(* CODESYS project process.library
   DefaultNamespace: KOSTAL.AF2024.Core.Process
   DocFormat: reStructuredText
   Description: Core Functionalities UTF16
   Author: Frank Dümpelmann
   Title: KOSTAL.AF2024.Core.Process
   Version: 1.0.999.1
   Company: KOSTAL GmbH & Co.KG
   Placeholder: KOSTAL.AF2024.Core.Process

Project tree, tasks and I/O mapping:
  libraries: KOSTAL.AF2024.Core.functionResponse, 1.0.0.0 (KOSTAL GmbH & Co.KG); KOSTAL.AF2024.Core.ListOf, 1.0.0.0 (KOSTAL GmbH & Co.KG); KOSTAL.AF2024.Core.Settings, 1.0.0.0 (KOSTAL GmbH & Co.KG); KOSTAL.AF2024.Core.StringTools, 1.0.0.0 (KOSTAL GmbH & Co.KG); KOSTAL.AF2024.Core.System, 1.0.0.0 (KOSTAL GmbH & Co.KG)
  _Global/
    E_/
      data type E_PROCESS_CONDITION_DEFAULT_PRIORITYLEVEL
  Condition/
    function block FB_processCondition [ST]: clear, CopyFrom, CopyTo, FB_init, getPriority, isActive, isError, isFail, isInfo, isMasterMessage, isMessage, isPass, isText, Message, Message_Owner, PriorityLevel_Error, PriorityLevel_Info, PriorityLevel_MasterMessage, PriorityLevel_Message, PriorityLevel_Text, setMessage, setMessageFail, setMessagePass
    interface I_processCondition: CopyTo, getPriority, isActive, isError, isFail, isInfo, isMasterMessage, isMessage, isPass, isText, Message, PriorityLevel_Error, PriorityLevel_Info, PriorityLevel_MasterMessage, PriorityLevel_Message, PriorityLevel_Text
    interface I_processCondition_CopyFrom: CopyFrom
    interface I_processCondition_Owner: clear, CopyFrom, CopyTo, getPriority, isActive, isError, isFail, isInfo, isMasterMessage, isMessage, isPass, isText, Message, Message_Owner, PriorityLevel_Error, PriorityLevel_Info, PriorityLevel_MasterMessage, PriorityLevel_Message, PriorityLevel_Text, setMessage, setMessageFail, setMessagePass
  DeviceState/
    interface I_T_deviceState: Fault, Off, On, Operational
    interface I_T_deviceState_Owner: ClearPlcState, Fault, Off, On, Operational
    function block T_deviceState [ST]: Clear, ClearPlcState, CopyFrom, CopyTo, Fault, Off, On, Operational
  Message/
    messageText/
      interface I_T_messageText: CopyTo, line_01, toString
      interface I_T_messageText_CopyFrom: CopyFrom
      interface I_T_messageText_Owner: clear, CopyFrom, CopyTo, line_01, toString
      function block T_messageText [ST]: clear, CopyFrom, CopyTo, line_01, toString
    messageText_2_lines/
      interface I_T_messageText_2_lines: line_02
      interface I_T_messageText_2_lines_Owner: line_02
      function block T_messageText_2_lines [ST]: clear, CopyFrom, line_02, toString
    messageText_3_lines/
      interface I_T_messageText_3_lines: line_03
      interface I_T_messageText_3_lines_Owner: line_03
      function block T_messageText_3_lines [ST]: clear, CopyFrom, line_03, toString
  PlcState/
    interface I_T_plcState: busy, CopyTo, description, fail, finish, pass, ready
    interface I_T_plcState_CopyFrom: CopyFrom
    interface I_T_plcState_Owner: busy, clear, CopyFrom, CopyTo, description, fail, finish, pass, ready
    function block T_plcState [ST]: busy, clear, CopyFrom, CopyTo, description, fail, finish, pass, ready
  ProcessMode/
    interface I_T_processMode: automatic, CopyTo, manual
    interface I_T_processMode_CopyFrom: CopyFrom
    interface I_T_processMode_Owner: automatic, clear, CopyFrom, CopyTo, manual
    function block T_processMode [ST]: automatic, clear, CopyFrom, CopyTo, manual
  Project Information/
    function F_GetCompany [ST]
    function F_GetTitle [ST]
    function F_GetVersion [ST]
  Step/
    GVL/
      global variables ProcessStep_GVL
    processStep/
      function block FB_processStep [ST]: actual, clear, CopyFrom, CopyTo, DEC, Header, INC, init, request, set, toggle
      interface I_processStep: actual, CopyTo, request, toggle
      interface I_processStep_CopyFrom: CopyFrom
      interface I_processStep_Owner: actual, clear, CopyFrom, CopyTo, DEC, Header, INC, init, request, set, toggle
    processStep_Control/
      StepMemory/
        ListOf/
          function block FB_ListOf_T_StepMemory [ST]: _get_I, _get_I_RO, _removePayLoad, _verifyMember, Add_DUT, Clear, CopyFrom, CopyTo, Delete_DUT, Get_I, Get_I_RO, MaxEntries, NumberOfMember
          interface I_ListOf_StepMemory: Add_DUT, Clear, CopyFrom, CopyTo, Delete_DUT, Get_I, Get_I_RO, MaxEntries, NumberOfMember
          interface I_ListOf_StepMemory_CopyFrom: CopyFrom
          interface I_ListOf_StepMemory_RO: CopyTo, Get_I_RO, MaxEntries, NumberOfMember
        interface I_T_StepMemory: Clear, CopyFrom, Actual, RegKey, Request
        interface I_T_StepMemory_CopyFrom: CopyFrom
        interface I_T_StepMemory_RO: CopyTo, Actual, RegKey, Request
        function block T_StepMemory [ST]: Clear, CopyFrom, CopyTo, Actual, RegKey, Request
      function block FB_ProcessStep_Control [ST]: FB_exit, FB_init, _DEC, _INC, _init, _set, _modeAutomatik, _backward, _forward, _modeManual, _addStep, _removeStep, _preset, DEC, INC, init, set, Control, clear, CopyFrom, Header, LinkManual, BackwardDone, Done, FromBackStep, LastUsedKey, StepMemory, StepMemory_RO, StepNumberHome, Condition, DisableBackward, JumpAddress, ManualWithCondition, mode
      interface I_ProcessStep_Control: BackwardDone, Done, FromBackStep, LastUsedKey, StepMemory_RO, StepNumberHome, Condition, DisableBackward, JumpAddress, ManualWithCondition, mode
      interface I_ProcessStep_Control_Owner: Control, Header, LinkManual, BackwardDone, Done, FromBackStep, LastUsedKey, StepMemory, StepMemory_RO, StepNumberHome, Condition, DisableBackward, JumpAddress, ManualWithCondition, mode
    processStep_Flow/
      function block FB_processStep_Flow [ST]: clear, Header, init, isActive, isCalledExternally, NotFound
      interface I_processStep_Flow: isCalledExternally, NotFound
      interface I_processStep_Flow_Owner: clear, Header, init, isActive, isCalledExternally, NotFound
  Version/
    global variables Global_Version
*)

// _Global/E_/E_PROCESS_CONDITION_DEFAULT_PRIORITYLEVEL
(*
Description
===========
| Levels of message priorities
| Intermediate values can be used to overrule other messages of the same level
| 1..999: INFORMATION - Display less important information (Color: grey)
| 1000..1999: TEXT_ONLY - To display information (Color: green)
| 2000..2999: MESSAGE - Order to the operator, e.g. 'Insert part' (Color: blue)
| 3000..3999: MASTERMESSAGE - Message to be displayed in upper HMI levels (Color: blue)
| 4000..4999: ERROR - Error message (Color: orange)

*)

{attribute 'qualified_only'}
TYPE E_PROCESS_CONDITION_DEFAULT_PRIORITYLEVEL :
(
	NONE 			:= 0,
	INFORMATION		:= 1,
	TEXT_ONLY		:= 1000,
	MESSAGE			:= 2000,
	MASTERMESSAGE	:= 3000,
	ERROR			:= 4000
);
END_TYPE

// Step/GVL/ProcessStep_GVL
{attribute 'qualified_only'}
VAR_GLOBAL CONSTANT
	PROCESS_STEP_INITIALIZE_STEP	: INT:= INT#32767; //INT[max] 16#7FFF;
END_VAR

// Version/Global_Version
{attribute 'TcGenerated'}
{attribute 'no-analysis'}
{attribute 'linkalways'}
// This function has been automatically generated from the project information.
VAR_GLOBAL CONSTANT
	{attribute 'const_non_replaced'}
	stLibVersion_KOSTAL_AF2024_Core_Process : ST_LibVersion := (iMajor := 1, iMinor := 0, iBuild := 999, iRevision := 1, nFlags := 1, sVersion := '1.0.999.1');
END_VAR

// Condition/FB_processCondition
(*

:Author: Frank Dümpelmann <f.duempelmann@kostal.com>
:Date: 2018-10-26

Function
========
| Data structure representing the status of users/stations 
| Used for communication to superior instances, e.g. HMI

Usage notes
===============
| Call method setMessage from User/Station to set Message Text and priority level
| Call methods is... from the superior instance to get the user's status 
| Read message text from property message 

Methods and Properties
======================
| See bottom of this document for a detailed description of each method or property
*)

{attribute 'enable_dynamic_creation'}
FUNCTION_BLOCK PUBLIC FB_processCondition IMPLEMENTS I_processCondition, I_processCondition_CopyFrom, I_processCondition_Owner

VAR
	_priority	: INT;	//Priority of message
	
	_message	: T_messageText_3_lines;
	
	_pass		: BOOL;
	_fail		: BOOL;
END_VAR

(*
Description
===========
| Clears existing message
*)

METHOD PUBLIC clear

_priority:= E_PROCESS_CONDITION_DEFAULT_PRIORITYLEVEL.NONE;

_message.clear();
_pass := _fail := false;
END_METHOD

METHOD PUBLIC CopyFrom : BOOL
VAR_INPUT
	IN	: KOSTAL_AF2024_Core_System.I_Interface;
END_VAR

VAR
	_obj		: I_processCondition;
	_obj2		: I_processCondition_Owner;
	_bFound	:	BOOL;
END_VAR

IF IN = 0 THEN	RETURN;	END_IF

clear();

//-----------------------------------------

_bFound:= __QUERYINTERFACE(IN, _obj);

IF _bFound AND_THEN _obj <> 0 THEN
	
	_priority:= _obj.getPriority();
	
	_message.CopyFrom(_obj.Message);
	
	_pass := _obj.isPass();
	_fail := _obj.isFail();
	
	
	CopyFrom:= TRUE;
	
	RETURN;
	
END_IF

//-----------------------------------------

_bFound:= __QUERYINTERFACE(IN, _obj2);

IF _bFound AND_THEN _obj2 <> 0 THEN
	
	_priority:= _obj2.getPriority();
	
	_message.CopyFrom(_obj2.Message);
	
	_pass := _obj2.isPass();
	_fail := _obj2.isFail();
	
	CopyFrom:= TRUE;

	RETURN;
	
END_IF
END_METHOD

METHOD PUBLIC CopyTo : BOOL
VAR_INPUT
	IN	:	I_processCondition_CopyFrom;
END_VAR

IF IN = 0 THEN	RETURN;	END_IF

CopyTo:= IN.CopyFrom(THIS^);
END_METHOD

(*
Description
===========
| To be called automatically!
*)
METHOD FB_init : BOOL
VAR_INPUT
	bInitRetains : BOOL; // if TRUE, the retain variables are initialized (warm start / cold start)
	bInCopyCode : BOOL;  // if TRUE, the instance afterwards gets moved into the copy code (online change)
END_VAR
//_infoPriorityLevel			:= E_PROCESS_CONDITION_DEFAULT_PRIORITYLEVEL.INFORMATION; 
//_textPriorityLevel			:= E_PROCESS_CONDITION_DEFAULT_PRIORITYLEVEL.TEXT_ONLY;		//define the priority level from which priority a message is an user relative text 
//_messagePriorityLevel		:= E_PROCESS_CONDITION_DEFAULT_PRIORITYLEVEL.MESSAGE;		//define the priority level from which priority a message is an user relative message 
//_masterMessagePriorityLevel	:= E_PROCESS_CONDITION_DEFAULT_PRIORITYLEVEL.MASTERMESSAGE;	//define the priority level from which priority a message is an user relative error 
//_errorPriorityLevel			:= E_PROCESS_CONDITION_DEFAULT_PRIORITYLEVEL.ERROR;			//define the priority level from which priority a message is an user relative error
END_METHOD

METHOD PUBLIC getPriority : INT
VAR_INPUT
END_VAR

getPriority:= _priority;
END_METHOD

(*
Description
===========
| Returns TRUE if the user has a text, message or error to display
*)

METHOD PUBLIC isActive : BOOL
VAR_INPUT
END_VAR

isActive:= _priority <> E_PROCESS_CONDITION_DEFAULT_PRIORITYLEVEL.NONE;
END_METHOD

(*
Description
===========
| Returns TRUE if the user has an error to display
*)
METHOD PUBLIC isError : BOOL
VAR_INPUT
END_VAR

isError:= _priority >= E_PROCESS_CONDITION_DEFAULT_PRIORITYLEVEL.ERROR;
END_METHOD

METHOD PUBLIC isFail : BOOL
VAR_INPUT
END_VAR
isFail := (isMessage() OR isMasterMessage()) AND _fail;
END_METHOD

(*
Description
===========
| Returns TRUE if the user has a message to display
*)
METHOD PUBLIC isInfo : BOOL
VAR_INPUT
END_VAR

isInfo:= (_priority >= E_PROCESS_CONDITION_DEFAULT_PRIORITYLEVEL.INFORMATION) AND (_priority < E_PROCESS_CONDITION_DEFAULT_PRIORITYLEVEL.TEXT_ONLY);
END_METHOD

(*
Description
===========
| Returns TRUE if the user has a master message to display
*)
METHOD PUBLIC isMasterMessage : BOOL
VAR_INPUT
END_VAR

isMasterMessage:= (_priority >= E_PROCESS_CONDITION_DEFAULT_PRIORITYLEVEL.MASTERMESSAGE) AND (_priority < E_PROCESS_CONDITION_DEFAULT_PRIORITYLEVEL.ERROR);
END_METHOD

(*
Description
===========
| Returns TRUE if the user has a message to display
*)
METHOD PUBLIC isMessage : BOOL
VAR_INPUT
END_VAR

isMessage:= (_priority >= E_PROCESS_CONDITION_DEFAULT_PRIORITYLEVEL.MESSAGE) AND (_priority < E_PROCESS_CONDITION_DEFAULT_PRIORITYLEVEL.MASTERMESSAGE);
END_METHOD

METHOD PUBLIC isPass : BOOL
VAR_INPUT
END_VAR
isPass := (isMessage() OR isMasterMessage()) AND _pass;
END_METHOD

(*
Description
===========
| Returns TRUE if the user has a text to display
*)
METHOD PUBLIC isText : BOOL

isText:= (_priority >= E_PROCESS_CONDITION_DEFAULT_PRIORITYLEVEL.TEXT_ONLY) AND (_priority < E_PROCESS_CONDITION_DEFAULT_PRIORITYLEVEL.MESSAGE);
END_METHOD

(*
Description
===========
| Message to display in three lines
*)

PROPERTY PUBLIC Message : I_T_messageText_3_lines
GET


Message := _message;
END_GET
END_PROPERTY

(*
Description
===========
| Message to display in three lines
*)

PROPERTY PUBLIC Message_Owner : I_T_messageText_3_lines_Owner
GET


Message_Owner := _message;
END_GET
END_PROPERTY

PROPERTY PUBLIC PriorityLevel_Error : INT
GET

PriorityLevel_Error := E_PROCESS_CONDITION_DEFAULT_PRIORITYLEVEL.ERROR;// _errorPriorityLevel;
END_GET
END_PROPERTY

PROPERTY PUBLIC PriorityLevel_Info : INT
GET

PriorityLevel_Info := E_PROCESS_CONDITION_DEFAULT_PRIORITYLEVEL.INFORMATION;
END_GET
END_PROPERTY

PROPERTY PUBLIC PriorityLevel_MasterMessage : INT
GET

PriorityLevel_MasterMessage := E_PROCESS_CONDITION_DEFAULT_PRIORITYLEVEL.MASTERMESSAGE;
END_GET
END_PROPERTY

PROPERTY PUBLIC PriorityLevel_Message : INT
GET

PriorityLevel_Message := E_PROCESS_CONDITION_DEFAULT_PRIORITYLEVEL.MESSAGE;
END_GET
END_PROPERTY

PROPERTY PUBLIC PriorityLevel_Text : INT
GET

PriorityLevel_Text := E_PROCESS_CONDITION_DEFAULT_PRIORITYLEVEL.TEXT_ONLY;
END_GET
END_PROPERTY

(*
Description
===========
| Sets message text and priority level for the user, in case the priority is higher than the existing message's priority 
| Existing messages with the same or lower priority are cleared
| Parameters:
| 	priority: INT - See E_PROCESS_CONDITION_DEFAULT_PRIORITYLEVEL for a detailed description
|	message: FB_messageText_3_lines - Content of the message
| Return value:
| 	FB_functionResponse: 
|		result: BOOL - Message ist set (no existing message with higher priority)
|		status: STRING(255) - Error description
*)

METHOD PUBLIC setMessage : KOSTAL_AF2024_Core_functionResponse.T_functionResponse

VAR_INPUT
	priority	: INT;
	message		: I_T_messageText_3_lines;
END_VAR
IF message = 0 THEN 
	setMessage.Status	:= "Message is invalid";
	setMessage.Success	:= FALSE;
	RETURN;	
END_IF

IF priority > _priority THEN
	setMessage.clear();
	_priority	:= priority;
	_message.CopyFrom(message);
	_pass := FALSE;
	_fail := FALSE;
	setMessage.Success	:= TRUE;

ELSE

	setMessage.Status	:= "actual priority is higher";
	setMessage.Success	:= FALSE;

END_IF
END_METHOD

(*
Description
===========
| Sets message text and priority level for the user, in case the priority is higher than the existing message's priority  
| Message is displayed as "Fail" (red) in WInHMI
| Existing messages with the same or lower priority are cleared
| Parameters:
| 	priority: INT - See E_PROCESS_CONDITION_DEFAULT_PRIORITYLEVEL for a detailed description
|	message: FB_messageText_3_lines - Content of the message
| Return value:
| 	FB_functionResponse: 
|		result: BOOL - Message ist set (no existing message with higher priority)
|		status: STRING(255) - Error description
*)

METHOD PUBLIC setMessageFail : KOSTAL_AF2024_Core_functionResponse.T_functionResponse

VAR_INPUT
	priority	: INT;
	message		: I_T_messageText_3_lines;
END_VAR
IF message = 0 THEN 
	setMessageFail.Status	:= "Message is invalid";
	setMessageFail.Success	:= FALSE;
	RETURN;	
END_IF

IF priority > _priority THEN
	setMessageFail.clear();
	_priority	:= priority;
	_message.CopyFrom(message);
	_pass := FALSE;
	_fail := TRUE;
	
	setMessageFail.Success	:= TRUE;

ELSE

	setMessageFail.Status	:= "actual priority is higher";
	setMessageFail.Success	:= FALSE;

END_IF
END_METHOD

(*
Description
===========
| Sets message text and priority level for the user, in case the priority is higher than the existing message's priority 
| Message is displayed as "Pass" (green) in WinHMI
| Existing messages with the same or lower priority are cleared
| Parameters:
| 	priority: INT - See E_PROCESS_CONDITION_DEFAULT_PRIORITYLEVEL for a detailed description
|	message: FB_messageText_3_lines - Content of the message
| Return value:
| 	FB_functionResponse: 
|		result: BOOL - Message ist set (no existing message with higher priority)
|		status: STRING(255) - Error description
*)

METHOD PUBLIC setMessagePass : KOSTAL_AF2024_Core_functionResponse.T_functionResponse

VAR_INPUT
	priority	: INT;
	message		: I_T_messageText_3_lines;
END_VAR
IF message = 0 THEN 
	setMessagePass.Status	:= "Message is invalid";
	setMessagePass.Success	:= FALSE;
	RETURN;	
END_IF

IF priority > _priority THEN
	setMessagePass.clear();
	_priority	:= priority;
	_message.CopyFrom(message);
	_pass := TRUE;
	_fail := FALSE;
	
	setMessagePass.Success	:= TRUE;

ELSE

	setMessagePass.Status	:= "actual priority is higher";
	setMessagePass.Success	:= FALSE;

END_IF
END_METHOD

END_FUNCTION_BLOCK

// Condition/I_processCondition
INTERFACE I_processCondition EXTENDS KOSTAL_AF2024_Core_System.I_Interface

METHOD PUBLIC CopyTo : BOOL
VAR_INPUT
	IN	:	I_processCondition_CopyFrom;
END_VAR
END_METHOD

METHOD PUBLIC getPriority : INT
VAR_INPUT
END_VAR
END_METHOD

(*
Description
===========
| Returns TRUE if the user has a text, message or error to display
*)

METHOD PUBLIC isActive : BOOL
VAR_INPUT
END_VAR
END_METHOD

(*
Description
===========
| Returns TRUE if the user has an error to display
*)
METHOD PUBLIC isError : BOOL
VAR_INPUT
END_VAR
END_METHOD

METHOD PUBLIC isFail : BOOL
VAR_INPUT
END_VAR
END_METHOD

(*
Description
===========
| Returns TRUE if the user has a message to display
*)
METHOD PUBLIC isInfo : BOOL
VAR_INPUT
END_VAR
END_METHOD

(*
Description
===========
| Returns TRUE if the user has a master message to display
*)
METHOD PUBLIC isMasterMessage : BOOL
VAR_INPUT
END_VAR
END_METHOD

(*
Description
===========
| Returns TRUE if the user has a message to display
*)
METHOD PUBLIC isMessage : BOOL
VAR_INPUT
END_VAR
END_METHOD

METHOD PUBLIC isPass : BOOL
VAR_INPUT
END_VAR
END_METHOD

(*
Description
===========
| Returns TRUE if the user has a text to display
*)
METHOD PUBLIC isText : BOOL
END_METHOD

(*
Description
===========
| Message to display in three lines
*)

PROPERTY PUBLIC Message : I_T_messageText_3_lines
GET
END_GET
END_PROPERTY

PROPERTY PUBLIC PriorityLevel_Error : INT
GET
END_GET
END_PROPERTY

PROPERTY PUBLIC PriorityLevel_Info : INT
GET
END_GET
END_PROPERTY

PROPERTY PUBLIC PriorityLevel_MasterMessage : INT
GET
END_GET
END_PROPERTY

PROPERTY PUBLIC PriorityLevel_Message : INT
GET
END_GET
END_PROPERTY

PROPERTY PUBLIC PriorityLevel_Text : INT
GET
END_GET
END_PROPERTY

END_INTERFACE

// Condition/I_processCondition_CopyFrom
INTERFACE I_processCondition_CopyFrom EXTENDS KOSTAL_AF2024_Core_System.I_Interface

METHOD PUBLIC CopyFrom : BOOL
VAR_INPUT
	IN	: KOSTAL_AF2024_Core_System.I_Interface;
END_VAR
END_METHOD

END_INTERFACE

// Message/messageText_3_lines/I_T_messageText_3_lines
INTERFACE I_T_messageText_3_lines EXTENDS I_T_messageText_2_lines

PROPERTY PUBLIC line_03 : KOSTAL_AF2024_Core_Settings.T_MaxString
GET
END_GET
END_PROPERTY

END_INTERFACE

// Message/messageText_2_lines/I_T_messageText_2_lines
INTERFACE I_T_messageText_2_lines EXTENDS I_T_messageText

PROPERTY PUBLIC line_02 : KOSTAL_AF2024_Core_Settings.T_MaxString
GET
END_GET
END_PROPERTY

END_INTERFACE

// Message/messageText/I_T_messageText
INTERFACE I_T_messageText EXTENDS KOSTAL_AF2024_Core_System.I_Interface

METHOD PUBLIC CopyTo : bool
VAR_INPUT
	IN	:	I_T_messageText_CopyFrom;
END_VAR
END_METHOD

PROPERTY PUBLIC line_01 : KOSTAL_AF2024_Core_Settings.T_MaxString
GET
END_GET
END_PROPERTY

METHOD PUBLIC toString : KOSTAL_AF2024_Core_Settings.T_MaxString
END_METHOD

END_INTERFACE

// Message/messageText/I_T_messageText_CopyFrom
INTERFACE I_T_messageText_CopyFrom

METHOD PUBLIC CopyFrom : BOOL
VAR_INPUT
	IN	: KOSTAL_AF2024_Core_System.I_Interface;
END_VAR
END_METHOD

END_INTERFACE

// Condition/I_processCondition_Owner
INTERFACE I_processCondition_Owner EXTENDS KOSTAL_AF2024_Core_System.I_Interface

(*
Description
===========
| Clears existing message
*)

METHOD PUBLIC clear
END_METHOD

METHOD PUBLIC CopyFrom : BOOL
VAR_INPUT
	IN	: KOSTAL_AF2024_Core_System.I_Interface;
END_VAR
END_METHOD

METHOD PUBLIC CopyTo : BOOL
VAR_INPUT
	IN	:	I_processCondition_CopyFrom;
END_VAR
END_METHOD

METHOD PUBLIC getPriority : INT
VAR_INPUT
END_VAR
END_METHOD

(*
Description
===========
| Returns TRUE if the user has a text, message or error to display
*)

METHOD PUBLIC isActive : BOOL
VAR_INPUT
END_VAR
END_METHOD

(*
Description
===========
| Returns TRUE if the user has an error to display
*)
METHOD PUBLIC isError : BOOL
VAR_INPUT
END_VAR
END_METHOD

METHOD PUBLIC isFail : BOOL
VAR_INPUT
END_VAR
END_METHOD

(*
Description
===========
| Returns TRUE if the user has a message to display
*)
METHOD PUBLIC isInfo : BOOL
VAR_INPUT
END_VAR
END_METHOD

(*
Description
===========
| Returns TRUE if the user has a master message to display
*)
METHOD PUBLIC isMasterMessage : BOOL
VAR_INPUT
END_VAR
END_METHOD

(*
Description
===========
| Returns TRUE if the user has a message to display
*)
METHOD PUBLIC isMessage : BOOL
VAR_INPUT
END_VAR
END_METHOD

METHOD PUBLIC isPass : BOOL
VAR_INPUT
END_VAR
END_METHOD

(*
Description
===========
| Returns TRUE if the user has a text to display
*)
METHOD PUBLIC isText : BOOL
END_METHOD

(*
Description
===========
| Message to display in three lines
*)

PROPERTY PUBLIC Message : I_T_messageText_3_lines
GET
END_GET
END_PROPERTY

(*
Description
===========
| Message to display in three lines
*)

PROPERTY PUBLIC Message_Owner : I_T_messageText_3_lines_Owner
GET
END_GET
END_PROPERTY

PROPERTY PUBLIC PriorityLevel_Error : INT
GET
END_GET
END_PROPERTY

PROPERTY PUBLIC PriorityLevel_Info : INT
GET
END_GET
END_PROPERTY

PROPERTY PUBLIC PriorityLevel_MasterMessage : INT
GET
END_GET
END_PROPERTY

PROPERTY PUBLIC PriorityLevel_Message : INT
GET
END_GET
END_PROPERTY

PROPERTY PUBLIC PriorityLevel_Text : INT
GET
END_GET
END_PROPERTY

(*
Description
===========
| Sets message text and priority level for the user, in case the priority is higher than the existing message's priority 
| Existing messages with the same or lower priority are cleared
| Parameters:
| 	priority: INT - See E_PROCESS_CONDITION_DEFAULT_PRIORITYLEVEL for a detailed description
|	message: FB_messageText_3_lines - Content of the message
| Return value:
| 	FB_functionResponse: 
|		result: BOOL - Message ist set (no existing message with higher priority)
|		status: STRING(255) - Error description
*)

METHOD PUBLIC setMessage : KOSTAL_AF2024_Core_functionResponse.T_functionResponse

VAR_INPUT
	priority	: INT;
	message		: I_T_messageText_3_lines;
END_VAR
END_METHOD

(*
Description
===========
| Sets message text and priority level for the user, in case the priority is higher than the existing message's priority 
| Message is displayed as "Fail" (red) in WInHMI
| Existing messages with the same or lower priority are cleared
| Parameters:
| 	priority: INT - See E_PROCESS_CONDITION_DEFAULT_PRIORITYLEVEL for a detailed description
|	message: FB_messageText_3_lines - Content of the message
| Return value:
| 	FB_functionResponse: 
|		result: BOOL - Message ist set (no existing message with higher priority)
|		status: STRING(255) - Error description
*)

METHOD PUBLIC setMessageFail : KOSTAL_AF2024_Core_functionResponse.T_functionResponse

VAR_INPUT
	priority	: INT;
	message		: I_T_messageText_3_lines;
END_VAR
END_METHOD

(*
Description
===========
| Sets message text and priority level for the user, in case the priority is higher than the existing message's priority  
| Message is displayed as "Pass" (green) in WinHMI
| Existing messages with the same or lower priority are cleared
| Parameters:
| 	priority: INT - See E_PROCESS_CONDITION_DEFAULT_PRIORITYLEVEL for a detailed description
|	message: FB_messageText_3_lines - Content of the message
| Return value:
| 	FB_functionResponse: 
|		result: BOOL - Message ist set (no existing message with higher priority)
|		status: STRING(255) - Error description
*)

METHOD PUBLIC setMessagePass : KOSTAL_AF2024_Core_functionResponse.T_functionResponse

VAR_INPUT
	priority	: INT;
	message		: I_T_messageText_3_lines;
END_VAR
END_METHOD

END_INTERFACE

// Message/messageText_3_lines/I_T_messageText_3_lines_Owner
INTERFACE I_T_messageText_3_lines_Owner EXTENDS I_T_messageText_2_lines_Owner

PROPERTY PUBLIC line_03 : KOSTAL_AF2024_Core_Settings.T_MaxString
GET
END_GET
SET
END_SET
END_PROPERTY

END_INTERFACE

// Message/messageText_2_lines/I_T_messageText_2_lines_Owner
INTERFACE I_T_messageText_2_lines_Owner EXTENDS I_T_messageText_Owner

PROPERTY PUBLIC line_02 : KOSTAL_AF2024_Core_Settings.T_MaxString
GET
END_GET
SET
END_SET
END_PROPERTY

END_INTERFACE

// Message/messageText/I_T_messageText_Owner
INTERFACE I_T_messageText_Owner EXTENDS KOSTAL_AF2024_Core_System.I_Interface

(*
Description
===========
| Clears existing text
*)

METHOD PUBLIC clear
VAR_INPUT
END_VAR
END_METHOD

METHOD PUBLIC CopyFrom : BOOL
VAR_INPUT
	IN	: KOSTAL_AF2024_Core_System.I_Interface;
END_VAR
END_METHOD

METHOD PUBLIC CopyTo : BOOL
VAR_INPUT
	IN	:	I_T_messageText_CopyFrom;
END_VAR
END_METHOD

PROPERTY PUBLIC line_01 : KOSTAL_AF2024_Core_Settings.T_MaxString
GET
END_GET
SET
END_SET
END_PROPERTY

METHOD PUBLIC toString : KOSTAL_AF2024_Core_Settings.T_MaxString
END_METHOD

END_INTERFACE

// Message/messageText_3_lines/T_messageText_3_lines
(*

:Author: Frank Dümpelmann <f.duempelmann@kostal.com>
:Date: 2018-10-26

Function
========
| Data type containing three lines of text
| To be used in HMI communication

Methods and Properties
======================
| Clear(): Clears existing text
| line_01, line_02, line_03: Lines of text
*)

{attribute 'enable_dynamic_creation'}
FUNCTION_BLOCK PUBLIC T_messageText_3_lines EXTENDS T_messageText_2_lines IMPLEMENTS I_T_messageText_3_lines, I_T_messageText_3_lines_Owner

VAR
	_line_03	: KOSTAL_AF2024_Core_Settings.T_MaxString;
END_VAR

(*
Description
===========
| Clears existing text
*)
METHOD PUBLIC clear
VAR_INPUT
END_VAR


SUPER^.clear();

_line_03:= "";
END_METHOD

METHOD PUBLIC CopyFrom : BOOL
VAR_INPUT
	IN	: KOSTAL_AF2024_Core_System.I_Interface;
END_VAR

VAR
	_obj		: I_T_messageText_3_lines;
	_obj2		: I_T_messageText_3_lines_Owner;
	_bFound: BOOL;
END_VAR

IF IN = 0 THEN	RETURN;	END_IF

clear();

//-----------------------------------------

_bFound := __QUERYINTERFACE(IN, _obj);
 
IF _bFound AND_THEN _obj <> 0 AND_THEN SUPER^.CopyFrom(IN) THEN

	_line_03	:= _obj.line_03;

	CopyFrom:= TRUE;

	RETURN;
	
END_IF

//-----------------------------------------

_bFound := __QUERYINTERFACE(IN, _obj2);
 
IF _bFound AND_THEN _obj2 <> 0 AND_THEN SUPER^.CopyFrom(IN) THEN

	_line_03	:= _obj2.line_03;
	CopyFrom:= TRUE;

	RETURN;	

END_IF
END_METHOD

PROPERTY PUBLIC line_03 : KOSTAL_AF2024_Core_Settings.T_MaxString
GET

line_03:= _line_03;
END_GET
SET

_line_03:= line_03;
END_SET
END_PROPERTY

METHOD PUBLIC toString : KOSTAL_AF2024_Core_Settings.T_MaxString

VAR
	_concat	: Kostal_AF2024_Core_StringTools.FB_Concat;	//KOSTAL_TC3_Components_Stringhandler.FB_CONCAT
END_VAR

_concat.clear();
_concat.addContent(SUPER^.toString());
_concat.addContent(";");
_concat.addContent(_line_03);

toString:= _concat.getResult();
END_METHOD

END_FUNCTION_BLOCK

// Message/messageText_2_lines/T_messageText_2_lines
(*

:Author: Frank Dümpelmann <f.duempelmann@kostal.com>
:Date: 2018-10-26

Function
========
| Data type containing two lines of text
| To be used in HMI communication

Methods and Properties
======================
| Clear(): Clears existing text
| line_01, line_02: Lines of text
*)

{attribute 'enable_dynamic_creation'}
FUNCTION_BLOCK PUBLIC T_messageText_2_lines EXTENDS T_messageText IMPLEMENTS I_T_messageText_2_lines, I_T_messageText_2_lines_Owner

VAR
	_line_02	: KOSTAL_AF2024_Core_Settings.T_MaxString;
END_VAR

(*
Description
===========
| Clears existing text
*)
METHOD PUBLIC clear
VAR_INPUT
END_VAR


SUPER^.clear();

_line_02:= "";
END_METHOD

METHOD PUBLIC CopyFrom : BOOL
VAR_INPUT
	IN	: KOSTAL_AF2024_Core_System.I_Interface;
END_VAR

VAR
	_obj		: I_T_messageText_2_lines;
	_obj2		: I_T_messageText_2_lines_Owner;
	_bFound	: BOOL;
END_VAR

IF IN = 0 THEN	RETURN;	END_IF

clear();

//-----------------------------------------

_bFound := __QUERYINTERFACE(IN, _obj);
 
IF _bFound AND_THEN _obj <> 0 AND_THEN SUPER^.CopyFrom(IN) THEN

	_line_02:= _obj.line_02;

	CopyFrom:= TRUE;

	RETURN;
	
END_IF

//-----------------------------------------

_bFound := __QUERYINTERFACE(IN, _obj2);
 
IF _bFound AND_THEN _obj2 <> 0 AND_THEN SUPER^.CopyFrom(IN) THEN

	_line_02:= _obj2.line_02;

	CopyFrom:= TRUE;

	RETURN;	

END_IF
END_METHOD

PROPERTY PUBLIC line_02 : KOSTAL_AF2024_Core_Settings.T_MaxString
GET

line_02:= _line_02;
END_GET
SET

_line_02:= line_02;
END_SET
END_PROPERTY

METHOD PUBLIC toString : KOSTAL_AF2024_Core_Settings.T_MaxString

VAR
	_concat	: Kostal_AF2024_Core_StringTools.FB_Concat;	//KOSTAL_TC3_Components_Stringhandler.FB_CONCAT
END_VAR

_concat.Clear();
_concat.addContent(SUPER^.toString());
_concat.addContent(";");
_concat.addContent(_line_02);

toString:= _concat.getResult();
END_METHOD

END_FUNCTION_BLOCK

// Message/messageText/T_messageText
(*

:Author: Frank Dümpelmann <f.duempelmann@kostal.com>
:Date: 2018-10-26

Function
========
| Data type containing one line of text
| To be used in HMI communication

Methods and Properties
======================
| Clear(): Clears existing text
| line_01: Line of text
*)

{attribute 'enable_dynamic_creation'}
FUNCTION_BLOCK PUBLIC T_messageText IMPLEMENTS I_T_messageText, I_T_messageText_CopyFrom, I_T_messageText_Owner

VAR
	_line_01	: KOSTAL_AF2024_Core_Settings.T_MaxString;
END_VAR

(*
Description
===========
| Clears existing text
*)

METHOD PUBLIC clear
VAR_INPUT
END_VAR

_line_01:= "";
END_METHOD

METHOD PUBLIC CopyFrom : BOOL
VAR_INPUT
	IN	: KOSTAL_AF2024_Core_System.I_Interface;
END_VAR

VAR
	_obj		: I_T_messageText;
	_obj2		: I_T_messageText_Owner;
	_bFound	:	BOOL;
END_VAR

IF IN = 0 THEN	RETURN;	END_IF

Clear();

//-----------------------------------------

_bFound:= __QUERYINTERFACE(IN, _obj);

IF _bFound AND_THEN _obj <> 0 THEN

	_line_01	:= _obj.line_01;

	CopyFrom:= TRUE;

	RETURN;	

END_IF
	
//-----------------------------------------

_bFound:= __QUERYINTERFACE(IN, _obj2);

IF _bFound AND_THEN _obj2 <> 0 THEN

	_line_01	:= _obj2.line_01;

	CopyFrom:= TRUE;

	RETURN;	

END_IF
END_METHOD

METHOD PUBLIC CopyTo : BOOL
VAR_INPUT
	IN	:	I_T_messageText_CopyFrom;
END_VAR

IF IN = 0 THEN	RETURN;	END_IF

CopyTo:= IN.CopyFrom(THIS^);
END_METHOD

PROPERTY PUBLIC line_01 : KOSTAL_AF2024_Core_Settings.T_MaxString
GET

line_01:= _line_01;
END_GET
SET

_line_01:= line_01;
END_SET
END_PROPERTY

METHOD PUBLIC toString : KOSTAL_AF2024_Core_Settings.T_MaxString

	
toString:= _line_01;
END_METHOD

END_FUNCTION_BLOCK

// DeviceState/I_T_deviceState
INTERFACE I_T_deviceState EXTENDS I_T_plcState

PROPERTY PUBLIC Fault : BOOL
GET
END_GET
END_PROPERTY

PROPERTY PUBLIC Off : BOOL
GET
END_GET
END_PROPERTY

PROPERTY PUBLIC On : BOOL
GET
END_GET
END_PROPERTY

PROPERTY PUBLIC Operational : BOOL
GET
END_GET
END_PROPERTY

END_INTERFACE

// PlcState/I_T_plcState
INTERFACE I_T_plcState EXTENDS KOSTAL_AF2024_Core_System.I_Interface

PROPERTY PUBLIC busy : BOOL
GET
END_GET
END_PROPERTY

METHOD PUBLIC CopyTo : BOOL
VAR_INPUT
	IN	:	I_T_plcState_CopyFrom;
END_VAR
END_METHOD

PROPERTY PUBLIC description : KOSTAL_AF2024_Core_Settings.T_MaxString
GET
END_GET
END_PROPERTY

PROPERTY PUBLIC fail : BOOL
GET
END_GET
END_PROPERTY

PROPERTY PUBLIC finish : BOOL
GET
END_GET
END_PROPERTY

PROPERTY PUBLIC pass : BOOL
GET
END_GET
END_PROPERTY

PROPERTY PUBLIC ready : BOOL
GET
END_GET
END_PROPERTY

END_INTERFACE

// PlcState/I_T_plcState_CopyFrom
INTERFACE I_T_plcState_CopyFrom EXTENDS KOSTAL_AF2024_Core_System.I_Interface

METHOD PUBLIC CopyFrom : BOOL
VAR_INPUT
	IN	: KOSTAL_AF2024_Core_System.I_Interface;
END_VAR
END_METHOD

END_INTERFACE

// DeviceState/I_T_deviceState_Owner
INTERFACE I_T_deviceState_Owner EXTENDS I_T_plcState_Owner

METHOD PUBLIC ClearPlcState
VAR_INPUT
END_VAR
END_METHOD

PROPERTY PUBLIC Fault : BOOL
GET
END_GET
SET
END_SET
END_PROPERTY

PROPERTY PUBLIC Off : BOOL
GET
END_GET
SET
END_SET
END_PROPERTY

PROPERTY PUBLIC On : BOOL
GET
END_GET
SET
END_SET
END_PROPERTY

PROPERTY PUBLIC Operational : BOOL
GET
END_GET
SET
END_SET
END_PROPERTY

END_INTERFACE

// PlcState/I_T_plcState_Owner
INTERFACE I_T_plcState_Owner EXTENDS KOSTAL_AF2024_Core_System.I_Interface

PROPERTY PUBLIC busy : BOOL
GET
END_GET
SET
END_SET
END_PROPERTY

METHOD PUBLIC clear
END_METHOD

METHOD PUBLIC CopyFrom : BOOL
VAR_INPUT
	IN	: KOSTAL_AF2024_Core_System.I_Interface;
END_VAR
END_METHOD

METHOD PUBLIC CopyTo : BOOL
VAR_INPUT
	IN	:	I_T_plcState_CopyFrom;
END_VAR
END_METHOD

PROPERTY PUBLIC description : KOSTAL_AF2024_Core_Settings.T_MaxString
GET
END_GET
SET
END_SET
END_PROPERTY

PROPERTY PUBLIC fail : BOOL
GET
END_GET
SET
END_SET
END_PROPERTY

PROPERTY PUBLIC finish : BOOL
GET
END_GET
SET
END_SET
END_PROPERTY

PROPERTY PUBLIC pass : BOOL
GET
END_GET
SET
END_SET
END_PROPERTY

PROPERTY PUBLIC ready : BOOL
GET
END_GET
SET
END_SET
END_PROPERTY

END_INTERFACE

// DeviceState/T_deviceState
(*

:Author: Frank Dümpelmann <f.duempelmann@kostal.com>
:Date: 2018-10-26

Function
========
Data type representing the process state of an item

Methods and Properties
======================
| Properties represent the possible process states (off, on, calibrate, ready, busy, finish)
| Methods setUnique_... set the corresponding state and clear the others
| Alternatively, states can be set independent of the others using the properties 
| Methods starting with an underline(_) are internally used and can be ignored by the user
*)
{attribute 'enable_dynamic_creation'}
FUNCTION_BLOCK PUBLIC T_deviceState EXTENDS T_plcState IMPLEMENTS I_T_deviceState, I_T_deviceState_Owner

VAR
	_off 					: BOOL;	//BOOL
	_on 					: BOOL;	//BOOL
	_operational	: BOOL;	//BOOL
	_fault				: BOOL;	//BOOL
END_VAR

METHOD PUBLIC Clear

SUPER^.Clear();

_off				 	:= FALSE;
_on 					:= FALSE;
_operational 	:= FALSE;
_fault				:= FALSE;
END_METHOD

METHOD PUBLIC ClearPlcState
VAR_INPUT
END_VAR

SUPER^.Clear();
END_METHOD

METHOD PUBLIC CopyFrom : BOOL
VAR_INPUT
	IN	: KOSTAL_AF2024_Core_System.I_Interface;
END_VAR

VAR
	_obj	: I_T_deviceState;
	_obj2	: I_T_deviceState_Owner;
	_bFound: BOOL;
END_VAR

IF IN = 0 THEN	RETURN;	END_IF

Clear();

//-----------------------------------------

_bFound := __QUERYINTERFACE(IN, _obj2);
 
IF _bFound AND_THEN _obj2 <> 0 AND_THEN SUPER^.CopyFrom(IN) THEN
	
	_off					:= _obj2.Off;
	_on						:= _obj2.on;
	_operational	:= _obj2.Operational;
	_fault				:= _obj2.Fault;

	CopyFrom:= TRUE;

	RETURN;
	
END_IF

//-----------------------------------------

_bFound := __QUERYINTERFACE(IN, _obj);
 
IF _bFound AND_THEN _obj <> 0 AND_THEN SUPER^.CopyFrom(IN) THEN
	
	_off					:= _obj.Off;
	_on						:= _obj.on;
	_operational	:= _obj.Operational;
	_fault				:= _obj.Fault;

	CopyFrom:= TRUE;

	RETURN;
	
END_IF
END_METHOD

METHOD PUBLIC CopyTo : BOOL
VAR_INPUT
	IN	:	I_T_plcState_CopyFrom;
END_VAR

IF IN = 0 THEN	RETURN;	END_IF

CopyTo:= IN.CopyFrom(THIS^);
END_METHOD

PROPERTY PUBLIC Fault : BOOL
GET

Fault:= _fault;
END_GET
SET

_fault:= Fault;
END_SET
END_PROPERTY

PROPERTY PUBLIC Off : BOOL
GET

off:= _off;
END_GET
SET

_off:= off;
END_SET
END_PROPERTY

PROPERTY PUBLIC On : BOOL
GET

On:= _on;
END_GET
SET

_on:= On;
END_SET
END_PROPERTY

PROPERTY PUBLIC Operational : BOOL
GET

Operational:= _operational;
END_GET
SET

_operational:= Operational;
END_SET
END_PROPERTY

END_FUNCTION_BLOCK

// PlcState/T_plcState
(*

:Author: Frank Dümpelmann <f.duempelmann@kostal.com>
:Date: 2018-10-26

Function
========
Data type representing the process state of an item

Methods and Properties
======================
| Properties represent the possible process states (off, on, calibrate, ready, busy, finish)
| Methods setUnique_... set the corresponding state and clear the others
| Alternatively, states can be set independent of the others using the properties 
| Methods starting with an underline(_) are internally used and can be ignored by the user
*)
{attribute 'enable_dynamic_creation'}
FUNCTION_BLOCK PUBLIC T_plcState IMPLEMENTS I_T_plcState, I_T_plcState_CopyFrom, I_T_plcState_Owner

VAR
	_ready 			: BOOL;	//BOOL
	_busy 			: BOOL;	//BOOL
	_finish 		: BOOL;	//BOOL
	_pass			: BOOL;
	_fail			: BOOL;
	_description	: KOSTAL_AF2024_Core_Settings.T_MaxString;
END_VAR

PROPERTY PUBLIC busy : BOOL
GET

busy:= _busy;
END_GET
SET

_busy:= busy;
END_SET
END_PROPERTY

METHOD PUBLIC clear

_busy		:= FALSE;
_finish		:= FALSE;

_ready		:= FALSE;
_pass		:= FALSE;
_fail		:= FALSE;

_description:= "";
END_METHOD

METHOD PUBLIC CopyFrom : BOOL
VAR_INPUT
	IN	: KOSTAL_AF2024_Core_System.I_Interface;
END_VAR


VAR
	_obj		: I_T_plcState;
	_obj2		: I_T_plcState_Owner;
	_bFound	:	BOOL;
END_VAR

IF IN = 0 THEN	RETURN;	END_IF

Clear();

//-----------------------------------------

_bFound:= __QUERYINTERFACE(IN, _obj);

IF _bFound AND_THEN _obj <> 0 THEN
	
	_ready				:= _obj.ready;
	_busy					:= _obj.busy;
	_finish				:= _obj.finish;
	_pass					:= _obj.pass;
	_fail					:= _obj.fail;
	_description 	:= _obj.description;

	CopyFrom:= TRUE;
	
	RETURN;

END_IF

//-----------------------------------------

_bFound:= __QUERYINTERFACE(IN, _obj2);

IF _bFound AND_THEN _obj2 <> 0 THEN
	
	_ready				:= _obj2.ready;
	_busy					:= _obj2.busy;
	_finish				:= _obj2.finish;
	_pass					:= _obj2.pass;
	_fail					:= _obj2.fail;
	_description 	:= _obj2.description;

	CopyFrom:= TRUE;

END_IF
END_METHOD

METHOD PUBLIC CopyTo : BOOL
VAR_INPUT
	IN	:	I_T_plcState_CopyFrom;
END_VAR

IF IN = 0 THEN	RETURN;	END_IF

CopyTo:= IN.CopyFrom(THIS^);
END_METHOD

PROPERTY PUBLIC description : KOSTAL_AF2024_Core_Settings.T_MaxString
GET

description:= _description;
END_GET
SET

_description:= description;
END_SET
END_PROPERTY

PROPERTY PUBLIC fail : BOOL
GET

fail:= _fail;
END_GET
SET

_fail:= fail;
END_SET
END_PROPERTY

PROPERTY PUBLIC finish : BOOL
GET

finish:= _finish;
END_GET
SET

_finish:= finish;
END_SET
END_PROPERTY

PROPERTY PUBLIC pass : BOOL
GET

pass:= _pass;
END_GET
SET

_pass:= pass;
END_SET
END_PROPERTY

PROPERTY PUBLIC ready : BOOL
GET

ready:= _ready;
END_GET
SET

_ready:= ready;
END_SET
END_PROPERTY

END_FUNCTION_BLOCK

// ProcessMode/I_T_processMode
INTERFACE I_T_processMode EXTENDS KOSTAL_AF2024_Core_System.I_Interface

PROPERTY PUBLIC automatic : BOOL
GET
END_GET
END_PROPERTY

METHOD PUBLIC CopyTo : bool
VAR_INPUT
	IN	:	I_T_processMode_CopyFrom;
END_VAR
END_METHOD

PROPERTY PUBLIC manual : BOOL
GET
END_GET
END_PROPERTY

END_INTERFACE

// ProcessMode/I_T_processMode_CopyFrom
INTERFACE I_T_processMode_CopyFrom EXTENDS KOSTAL_AF2024_Core_System.I_Interface

METHOD PUBLIC CopyFrom : BOOL
VAR_INPUT 
	IN	: KOSTAL_AF2024_Core_System.I_Interface;
END_VAR
END_METHOD

END_INTERFACE

// ProcessMode/I_T_processMode_Owner
INTERFACE I_T_processMode_Owner EXTENDS KOSTAL_AF2024_Core_System.I_Interface

PROPERTY PUBLIC automatic : BOOL
GET
END_GET
SET
END_SET
END_PROPERTY

METHOD PUBLIC clear
END_METHOD

METHOD PUBLIC CopyFrom : BOOL
VAR_INPUT
	IN	: KOSTAL_AF2024_Core_System.I_Interface;
END_VAR
END_METHOD

METHOD PUBLIC CopyTo : BOOL
VAR_INPUT
	IN	:	I_T_processMode_CopyFrom;
END_VAR
END_METHOD

PROPERTY PUBLIC manual : BOOL
GET
END_GET
SET
END_SET
END_PROPERTY

END_INTERFACE

// ProcessMode/T_processMode
(*

:Author: Frank Dümpelmann <f.duempelmann@kostal.com>
:Date: 2018-10-26

Function
========
Data type representing the manual/automatic mode of an item
*)
{attribute 'enable_dynamic_creation'}
FUNCTION_BLOCK PUBLIC T_processMode IMPLEMENTS I_T_processMode, I_T_processMode_CopyFrom, I_T_processMode_Owner

VAR
	_automatic	: BOOL;	//Release Automatic Functions
	_manual		: BOOL;	//Release Manual Functions	
END_VAR

PROPERTY PUBLIC automatic : BOOL
GET

automatic:= _automatic;
END_GET
SET

_automatic:= automatic;
END_SET
END_PROPERTY

METHOD PUBLIC clear

_automatic:= FALSE;
_manual		:= FALSE;
END_METHOD

METHOD PUBLIC CopyFrom : BOOL
VAR_INPUT
	IN	: KOSTAL_AF2024_Core_System.I_Interface;
END_VAR

VAR
	_obj		: I_T_processMode_Owner;
	_obj2		: I_T_processMode;
	_bFound	:	BOOL;
END_VAR

IF IN = 0 THEN	RETURN;	END_IF

Clear();

//-----------------------------------------

_bFound:= __QUERYINTERFACE(IN, _obj);

IF _bFound AND_THEN _obj <> 0 THEN

	_automatic	:= _obj.automatic;
	_manual			:= _obj.manual;


	CopyFrom:= TRUE;

	RETURN;
	
END_IF

//-----------------------------------------
	
_bFound:= __QUERYINTERFACE(IN, _obj2);

IF _bFound AND_THEN _obj2 <> 0 THEN

	_automatic	:= _obj2.automatic;
	_manual			:= _obj2.manual;

	CopyFrom:= TRUE;

	RETURN;
	
END_IF
END_METHOD

METHOD PUBLIC CopyTo : BOOL
VAR_INPUT
	IN	:	I_T_processMode_CopyFrom;
END_VAR

IF IN = 0 THEN	RETURN;	END_IF

CopyTo:= IN.CopyFrom(THIS^);
END_METHOD

PROPERTY PUBLIC manual : BOOL
GET

manual:= _manual;
END_GET
SET

_manual:= manual;
END_SET
END_PROPERTY

END_FUNCTION_BLOCK

// Project Information/F_GetCompany
// This function has been automatically generated from the project information.
{attribute 'signature_flag' := '1073741824'}
{attribute 'TcGenerated'}
{attribute 'no-analysis'}
FUNCTION F_GetCompany : WSTRING
VAR_INPUT
	
END_VAR

F_GetCompany := "KOSTAL GmbH & Co.KG";

END_FUNCTION

// Project Information/F_GetTitle
// This function has been automatically generated from the project information.
{attribute 'signature_flag' := '1073741824'}
{attribute 'TcGenerated'}
{attribute 'no-analysis'}
FUNCTION F_GetTitle : WSTRING
VAR_INPUT
	
END_VAR

F_GetTitle := "KOSTAL.AF2024.Core.Process";

END_FUNCTION

// Project Information/F_GetVersion
// This function has been automatically generated from the project information.
{attribute 'signature_flag' := '1073741824'}
{attribute 'TcGenerated'}
{attribute 'no-analysis'}
FUNCTION F_GetVersion : ST_LibVersion
VAR_INPUT
	
END_VAR

F_GetVersion.iMajor := 1;
F_GetVersion.iMinor := 0;
F_GetVersion.iBuild := 999;
F_GetVersion.iRevision := 1;
F_GetVersion.sVersion := '1.0.999.1';
F_GetVersion.nFlags := 1;

END_FUNCTION

// Step/processStep/FB_processStep
(*

:Author: Frank Dümpelmann <f.duempelmann@kostal.com>
:Date: 2018-10-26

Function
========
| Data structure representing a step sequence or state machine
| All changes are applied when the method Header() is called
| For the main step sequence of a station, use FB_ProcessStep_Control (implementig manual/automatic,...)

Methods and Properties
======================
| See bottom of this document for a detailed description of each method or property
| Methods starting with an underline(_) are internally used and can be ignored by the user

Usage sample:
=============

.. code:: 

	PROGRAM MAIN
	VAR
		_step : FB_processStep;
		_reset : BOOL := TRUE;
		_test1: BOOL;	
		_test2: INT;
		_test3: BOOL;
		_test4: BOOL;
	END_VAR
	
	IF _reset THEN
		_step.init();	//Init
		_reset := FALSE;
	END_IF
	
	_step.Header(); //Call before step sequence
	
	CASE _step.actual OF 
		0: 	IF (_test1) THEN
				_step.INC();	//Increase by one
			END_IF
		1: 	IF (_test2 > 1) THEN
				_step.request := 3;	//Set requested number directly
			ELSE
				_step.request := 4;	
			END_IF
		3: 	IF _test4 THEN
				_step.set(5);	//Set Method
			END_IF
			
		4: 	IF _test3 THEN
			_step.DEC();		//Decrease by one
			END_IF
		5: _reset := true;
	END_CASE
	
	IF _step.toggle THEN
	_toggleCounter := _toggleCounter+1;
	END_IF

*)

{attribute 'enable_dynamic_creation'}
FUNCTION_BLOCK FB_processStep IMPLEMENTS I_processStep, I_processStep_CopyFrom, I_processStep_Owner

VAR
	_actual						: INT ;	//Actual Step Number
	_request					: INT;	//Requested Step Number
	_toggle						: BOOL;	//TRUE if actual Step Number is actualized with the requested
END_VAR

(*
Description
===========
| Actual step number
*)
PROPERTY PUBLIC actual : INT
GET

actual:= _actual;
END_GET
END_PROPERTY

METHOD PUBLIC clear

_actual		:= 0;
_request	:= 0;
_toggle		:= FALSE;
END_METHOD

METHOD PUBLIC CopyFrom : BOOL
VAR_INPUT
	IN	: KOSTAL_AF2024_Core_System.I_Interface;
END_VAR

VAR
	_obj		:	I_processStep;
	_obj2		:	I_processStep_Owner;
	_bFound	: BOOL;
END_VAR

IF IN = 0 THEN	RETURN;	END_IF

clear();

//-----------------------------------------

_bFound:= __QUERYINTERFACE(IN, _obj);

IF _bFound AND_THEN _obj <> 0 THEN

	_actual		:= _obj.actual;
	_request	:= _obj.request;
	_toggle		:= _obj.toggle;

	CopyFrom	:= TRUE;

	RETURN;

END_IF


//-----------------------------------------

_bFound:= __QUERYINTERFACE(IN, _obj2);

IF _bFound AND_THEN _obj2 <> 0 THEN

	_actual		:= _obj2.actual;
	_request	:= _obj2.request;
	_toggle		:= _obj2.toggle;

	CopyFrom	:= TRUE;

	RETURN;

END_IF
END_METHOD

METHOD PUBLIC CopyTo : BOOL
VAR_INPUT
	IN	:	I_processStep_CopyFrom;
END_VAR

IF IN = 0 THEN	RETURN;	END_IF

CopyTo:= IN.CopyFrom(THIS^);
END_METHOD

(*
Description
===========
| Decrease step number by one (will be set with the next call of Header()
*)
METHOD DEC : KOSTAL_AF2024_Core_functionResponse.T_functionResponse
VAR_INPUT
END_VAR

IF (_actual - 1) >  _actual THEN

	DEC.status	:= "Overflow";
	DEC.success	:= FALSE;

ELSE

	_request:= _actual - 1;

	DEC.status	:= "";
	DEC.success	:= TRUE;
	
END_IF
END_METHOD

(*
Description
===========
| Apply changes in step sequence
| Call before or after the step sequence (see usage sample)
*)
METHOD PUBLIC Header
VAR_INPUT
END_VAR
_toggle:= _actual <> _request;
_actual := _request;
END_METHOD

(*
Description
===========
| Increase step number by one (will be set with the next call of Header()
*)
METHOD INC : KOSTAL_AF2024_Core_functionResponse.T_functionResponse
VAR_INPUT
END_VAR


IF (_actual + 1) <  _actual THEN

	INC.Status	:= "Overflow";
	INC.Success	:= FALSE;

ELSE

	_request:= _actual + 1;

	INC.Status	:= "";
	INC.Success	:= TRUE;
	
END_IF
END_METHOD

(*
Description
===========
| Reset step sequence to 0
*)
METHOD PUBLIC init


_actual		:= ProcessStep_GVL.PROCESS_STEP_INITIALIZE_STEP;	//UINT_TO_INT(16#FFFF);
_request	:= 0;
_toggle		:= TRUE;
END_METHOD

(*
Description
===========
| Requested step number (will be set with the next call of Header()
*)
PROPERTY PUBLIC request : INT
GET

request:= _request;
END_GET
END_PROPERTY

(*
Description
===========
| Select step number (will be set with the next call of Header()
| Same function as property request
| Parameters:
| 	request: INT - step number to go to
*)
METHOD PUBLIC set

VAR_INPUT
	request	: INT;	//INT
END_VAR


_request:= request;
END_METHOD

(*
Description
===========
| Toggle signal for initialzation purposes
| Is set TRUE when Header() was called and the step number changed
| Is reset FALSE with the next call of Header() without changing step number
*)

PROPERTY PUBLIC toggle : BOOL
GET

toggle:= _toggle;
END_GET
END_PROPERTY

END_FUNCTION_BLOCK

// Step/processStep_Control/FB_ProcessStep_Control
(*

:Author: Frank Dümpelmann <f.duempelmann@kostal.com>
:Date: 2018-10-26

Function
========
| Function block implementing the main step sequence of a station
| Variable step numbers, stepping forward and backward
| Feedback of successful step change
| Selection of manual or automatic stepping


Usage notes
===============
| Call method Header() before the step sequence
| Call method Control() at the end of each step to check the stepping condition 

Methods and Properties
======================
| See bottom of this document for a detailed description of each method or property
| Methods starting with an underline(_) are internally used and can be ignored by the user

*)

{attribute 'enable_dynamic_creation'}
FUNCTION_BLOCK PUBLIC FB_ProcessStep_Control EXTENDS FB_processStep IMPLEMENTS I_ProcessStep_Control, I_ProcessStep_Control_Owner

VAR

	_mode	: T_processMode;	//ST_ProcessMode

	_condition						: BOOL;	//BOOL
	_manualWithCondition	: BOOL;	//BOOL
	_manualForward				: BOOL;	//BOOL
	_manualBackward				: BOOL;	//BOOL
	_disableBackward			: BOOL; //TRUE > denies a DEC operation

	_jumpAddress					:	INT;	//INT

	_called				: BOOL;	//TRUE if one of the public methods is called in this cycle
	_done					: BOOL;	//TRUE on each event
	_backwardDone	: BOOL;	//TRUE if use DEC()
	_FromBackStep	: BOOL;	//Step was selected via a DEC method.


	_lastUsedKey	: ULINT;//Last Key used in _addStep or _removeStep

	{region 'StepMemory'}
		//defines the step number above which a StepMemory is created and from which a manual cycle is accepted back.
		_StepNumberHome	: INT:= ProcessStep_GVL.PROCESS_STEP_INITIALIZE_STEP;
	
		//Memory of the steps executed in this cycle.
		_stepMemory	: FB_ListOf_T_StepMemory;
	{endregion}

	_response	:	KOSTAL_AF2024_Core_functionResponse.T_functionResponse;
	
END_VAR

METHOD FB_exit : BOOL
VAR_INPUT
	bInCopyCode : BOOL; // if TRUE, the exit method is called for exiting an instance that is copied afterwards (online change).
END_VAR

_stepMemory.Clear();
END_METHOD

METHOD FB_init : BOOL
VAR_INPUT
	bInitRetains : BOOL; // if TRUE, the retain variables are initialized (warm start / cold start)
	bInCopyCode : BOOL;  // if TRUE, the instance afterwards gets moved into the copy code (online change)
END_VAR

_stepMemory.Clear();
END_METHOD

(*
Description
===========
| Decrease step number by one (will be set with the next call of Header()
*)
METHOD PROTECTED _DEC : KOSTAL_AF2024_Core_functionResponse.T_functionResponse
VAR
	_Mem	: T_StepMemory;
	_IMem	: I_T_StepMemory;
END_VAR

_preset();

_DEC:= SUPER^.DEC();

IF NOT _DEC.success	THEN RETURN;	END_IF

IF _request > _StepNumberHome	THEN _addStep();	END_IF

_done			:= TRUE;
//_decDone	:= TRUE;
END_METHOD

(*
Description
===========
| Increase step number by one (will be set with the next call of Header()
*)
METHOD PROTECTED _INC : KOSTAL_AF2024_Core_functionResponse.T_functionResponse
VAR_INPUT
END_VAR

_preset();

_INC:= SUPER^.INC();

IF NOT _INC.success	THEN RETURN;	END_IF

IF _request > _StepNumberHome	THEN _addStep();	END_IF

_done			:= TRUE;
//_incDone	:= TRUE;
END_METHOD

(*
Description
===========
| Reset step sequence to 0
*)
METHOD PROTECTED  _init

_preset();

SUPER^.init();

_stepMemory.Clear();

_done			:= TRUE;
END_METHOD

(*
Description
===========
| Select step number (will be set with the next call of Header()
| Same function as property request
| Parameters:
| 	request: INT - step number to go to
*)
METHOD PROTECTED  _set

VAR_INPUT
	request	: INT;	//INT
END_VAR

_preset();

SUPER^.set(request);

IF _actual <> _request AND_THEN _request > _StepNumberHome THEN	_addStep();	END_IF

_done			:= TRUE;
//_setDone	:= TRUE;
END_METHOD

METHOD PROTECTED _modeAutomatik : KOSTAL_AF2024_Core_functionResponse.T_functionResponse


IF _condition THEN

	_condition:= FALSE;
	
	IF _jumpAddress <> 0 THEN

		_set(_jumpAddress);
		
		_modeAutomatik.Status	:= "";
		_modeAutomatik.Success:= TRUE;
		
	ELSE
		
		_modeAutomatik:= _INC();
	
	END_IF

ELSE
	
	_modeAutomatik.Status	:= "Wait for condition";
	_modeAutomatik.Success:= FALSE;

END_IF
END_METHOD

(*
Description
===========
| Decrease step number by one (will be set with the next call of Header()
*)
METHOD PROTECTED _backward : KOSTAL_AF2024_Core_functionResponse.T_functionResponse
VAR
	_Mem	: T_StepMemory;
	_IMem	: I_T_StepMemory;
END_VAR

IF _disableBackward THEN 

	_backward.success:= FALSE;
	_backward.status:= "Backward disabled";

	RETURN;

END_IF

_preset();

IF NOT _stepMemory.Get_I(_stepMemory.NumberOfMember, _IMem, _response)	THEN _backward.CopyFrom(_response); RETURN;	END_IF
 
IF _IMem.Request <> _actual THEN _backward.success:= FALSE;	_backward.status:= "No matching step element found";	RETURN;	END_IF

SUPER^.set(_IMem.Actual);

_removeStep();	

_backward.success:= TRUE;
_backward.status:= "_backward successfull";

_done					:= TRUE;
_backwardDone	:= TRUE;
_FromBackStep	:= TRUE;
END_METHOD

METHOD PROTECTED _forward : KOSTAL_AF2024_Core_functionResponse.T_functionResponse

IF _jumpAddress <> 0 THEN

	_set(_jumpAddress);

	_Forward.Status		:= "";
	_Forward.Success	:= TRUE;

ELSE

		_Forward:= _INC();

END_IF
END_METHOD

METHOD PROTECTED _modeManual : KOSTAL_AF2024_Core_functionResponse.T_functionResponse


IF NOT _manualWithCondition OR _condition THEN

	_condition:= FALSE;
	
	IF _manualForward THEN

		_modeManual:= _forward();
		
		_manualForward	:= FALSE;

//		IF _modeManual.Success THEN
//			_forwardDone		:= TRUE;	
//		END_IF

	ELSIF _manualBackward THEN
		
		_modeManual:=  _backward();

		_manualBackward	:= FALSE;	
		
		IF _modeManual.Success THEN	
			_backwardDone		:= TRUE;	
		END_IF

	ELSE

	_modeManual.Status:= "Wait for manual request";
	_modeManual.Success:= FALSE;
		
	END_IF


ELSE
		
	_modeManual.Status:= "Wait for condition";
	_modeManual.Success:= FALSE;

END_IF
END_METHOD

METHOD PROTECTED _addStep : BOOL

VAR
	_Mem	: T_StepMemory;
	_iStepMem	: I_T_StepMemory_RO;
END_VAR

_Mem.Actual:= _actual;
_Mem.Request:= _request;

_addStep:= _StepMemory.Add_DUT(_Mem, 0);

IF 				_addStep 
AND_THEN	_StepMemory.Get_I_RO(_StepMemory.NumberOfMember, _iStepMem, 0)	
AND_THEN	_iStepMem <> 0
THEN			_lastUsedKey:= _iStepMem.RegKey;
END_IF
END_METHOD

METHOD PROTECTED _removeStep : BOOL
VAR
	_iStepMem	: I_T_StepMemory_RO;
END_VAR

IF 				_StepMemory.Get_I_RO(_StepMemory.NumberOfMember, _iStepMem, 0)	
AND_THEN	_iStepMem <> 0
THEN			_lastUsedKey:= _iStepMem.RegKey;
END_IF

_removeStep:= _StepMemory.Delete_DUT(_StepMemory.NumberOfMember, 0);
END_METHOD

METHOD PROTECTED _preset : BOOL

_jumpAddress					:= 0;
_condition						:= FALSE;
_FromBackStep					:= FALSE;
_disableBackward			:= FALSE;
_manualWithCondition	:= FALSE;
END_METHOD

(*
Description
===========
| Decrease step number by one (will be set with the next call of Header()
*)
METHOD DEC : KOSTAL_AF2024_Core_functionResponse.T_functionResponse
VAR
	_Mem	: T_StepMemory;
	_IMem	: I_T_StepMemory;
END_VAR

IF _called	THEN	RETURN;	END_IF
_called:= TRUE;

DEC:= _DEC();
END_METHOD

(*
Description
===========
| Increase step number by one (will be set with the next call of Header()
*)
METHOD INC : KOSTAL_AF2024_Core_functionResponse.T_functionResponse
VAR_INPUT
END_VAR

IF _called	THEN	RETURN;	END_IF
_called:= TRUE;

INC:= _INC();
END_METHOD

(*
Description
===========
| Reset step sequence to 0
*)
METHOD PUBLIC init

_init();
END_METHOD

(*
Description
===========
| Select step number (will be set with the next call of Header()
| Same function as property request
| Parameters:
| 	request: INT - step number to go to
*)
METHOD PUBLIC set

VAR_INPUT
	request	: INT;	//INT
END_VAR

IF _called	THEN	RETURN;	END_IF
_called:= TRUE;

_set(request);
END_METHOD

(*
Description
===========
| Select next step number dependent of Condition and JumpAddress
*)

METHOD PUBLIC Control : KOSTAL_AF2024_Core_functionResponse.T_functionResponse

IF _called	THEN	RETURN;	END_IF


IF _mode.Automatic THEN
	
	Control := _modeAutomatik();
	IF Control.success THEN _called:= TRUE;	END_IF
	
ELSIF _mode.Manual THEN

	Control := _modeManual();
	IF Control.success THEN _called:= TRUE;	END_IF

ELSE

	Control.Status:= "no mode detected";
	Control.Success:= FALSE;

END_IF
END_METHOD

METHOD PUBLIC clear

SUPER^.clear();

_condition						:= FALSE;
_done									:= FALSE;
_backwardDone					:= FALSE;
_manualWithCondition	:= FALSE;

_jumpAddress					:= 0;

_mode.clear();

_stepMemory.Clear();
END_METHOD

METHOD PUBLIC CopyFrom : BOOL
VAR_INPUT
	IN	: KOSTAL_AF2024_Core_System.I_Interface;
END_VAR

VAR
	_obj		: I_ProcessStep_Control;
	_obj2		: I_ProcessStep_Control_Owner;
	_bFound	: BOOL;
END_VAR

IF IN = 0 THEN RETURN;	END_IF

clear();

//-----------------------------------------

_bFound:= __QUERYINTERFACE(IN, _obj);

IF _bFound AND_THEN _obj <> 0 AND_THEN SUPER^.CopyFrom(IN) THEN
	
	_condition						:= _obj.Condition;
	
	_done									:= _obj.Done;
	_backwardDone					:= _obj.BackwardDone;
	_jumpAddress					:= _obj.JumpAddress;
	_manualWithCondition	:= _obj.ManualWithCondition;
	_mode									:= _obj.mode;
	
	_stepMemory.CopyFrom(_obj.StepMemory_RO);

	CopyFrom:= TRUE;

	RETURN;
	
END_IF


//-----------------------------------------

_bFound:= __QUERYINTERFACE(IN, _obj2);

IF _bFound AND_THEN _obj2 <> 0 AND_THEN SUPER^.CopyFrom(IN) THEN
	
	_condition						:= _obj2.Condition;
	
	_done									:= _obj2.Done;
	_backwardDone					:= _obj2.BackwardDone;
	_jumpAddress					:= _obj2.JumpAddress;
	_manualWithCondition	:= _obj2.ManualWithCondition;
	_mode									:= _obj2.mode;
	
	_stepMemory.CopyFrom(_obj2.StepMemory_RO);

	CopyFrom:= TRUE;

	RETURN;
	
END_IF
END_METHOD

(*
Description
===========
| Apply changes in step sequence
| Call before the step sequence (see usage sample)
*)
METHOD PUBLIC Header


super^.Header();

IF _toggle AND_THEN (_actual <= _StepNumberHome) AND_THEN (_stepMemory.NumberOfMember > 0) THEN	_stepMemory.Clear();	END_IF

_called				:= FALSE;
_done					:= FALSE;

//_incDone			:= FALSE;
//_decDone			:= FALSE;
//_setDone			:= FALSE;
//_initDone			:= FALSE;

_backwardDone	:= FALSE;
//_forwardDone	:= FALSE;
END_METHOD

//It is mandatory to link the parameters exclusively with pulses. 
METHOD PUBLIC LinkManual
VAR_INPUT
	Forward		: BOOL;	//Pulse one step forward in the step chain 
	Backward	: BOOL;	//Pulse one step backwards in the step chain
END_VAR

_manualForward	:= Forward;
_manualBackward	:= Backward;
END_METHOD

(*
Description
===========
| Step change backward was successful - Use e.g. to reset requests
| Attention: Variable is reset with next call of Header()
*)
PROPERTY PUBLIC BackwardDone : BOOL
GET

IF _actual <> _request THEN	BackwardDone:= _backwardDone;	
ELSE												BackwardDone:= FALSE;
END_IF
END_GET
END_PROPERTY

(*
Description
===========
| Step change was successful - Use e.g. to reset requests
| Attention: Variable is reset with next call of Header()
*)
PROPERTY PUBLIC Done : BOOL
GET

IF _actual <> _request THEN	Done:= _done;	
ELSE												Done:= FALSE;
END_IF
END_GET
END_PROPERTY

PROPERTY PUBLIC FromBackStep : BOOL
GET

FromBackStep:= _FromBackStep;
END_GET
END_PROPERTY

PROPERTY PUBLIC LastUsedKey : ULINT
GET

LastUsedKey:= _lastUsedKey;
END_GET
END_PROPERTY

PROPERTY PUBLIC StepMemory : I_ListOf_StepMemory
GET

StepMemory:= _stepMemory;
END_GET
END_PROPERTY

PROPERTY PUBLIC StepMemory_RO : I_ListOf_StepMemory_RO
GET

StepMemory_RO:= _stepMemory;
END_GET
END_PROPERTY

PROPERTY PUBLIC StepNumberHome : INT
GET

StepNumberHome:= _StepNumberHome;
END_GET
SET

_StepNumberHome:= StepNumberHome;
END_SET
END_PROPERTY

(*
Description
===========
| Condition to switch to the next step in automatic mode (also in manual mode if "ManualWithCondition" is TRUE) 
*)

PROPERTY PUBLIC Condition : BOOL
GET

Condition:= _condition;
END_GET
SET

_condition:= Condition;
END_SET
END_PROPERTY

PROPERTY PUBLIC DisableBackward : BOOL
GET

DisableBackward:= _disableBackward;
END_GET
SET

_disableBackward:= DisableBackward;
END_SET
END_PROPERTY

(*
Description
===========
| Step number to go to next
| 0 = subsequent step
*)
PROPERTY PUBLIC JumpAddress : INT
GET


JumpAddress:= _jumpAddress;
END_GET
SET

_jumpAddress:= JumpAddress;
END_SET
END_PROPERTY

(*
Description
===========
| If TRUE, property "Condition" is also active in manual mode
*)
PROPERTY PUBLIC ManualWithCondition : BOOL
GET

ManualWithCondition:= _manualWithCondition;
END_GET
SET

_manualWithCondition:= ManualWithCondition;
END_SET
END_PROPERTY

(*
Description
===========
| automatic: Control automatically jumps to the next step if Condition is TRUE
| manual: Input ManualForward must be pulsed TRUE to go to the next step
*)
PROPERTY PUBLIC mode : REFERENCE to T_processMode
GET

mode REF= _mode;
END_GET
SET

_mode := mode;
END_SET
END_PROPERTY

END_FUNCTION_BLOCK

// Step/processStep_Control/I_ProcessStep_Control
(*

:Author: Martin Hundt <m.hundt@kostal.com>
:Date: 2019-04-18

Function
========
Interface to link current state/content from FB_ProcessStep_Control to other components which analyse the step sequence internally (e.g. FB_Cylinder_Controlled)
*)
INTERFACE I_ProcessStep_Control EXTENDS I_processStep

(*
Description
===========
| Step change backward was successful - Use e.g. to reset requests
| Attention: Variable is reset with next call of Header()
*)
PROPERTY PUBLIC BackwardDone : BOOL
GET
END_GET
END_PROPERTY

(*
Description
===========
| Step change was successful - Use e.g. to reset requests
| Attention: Variable is reset with next call of Header()
*)
PROPERTY PUBLIC Done : BOOL
GET
END_GET
END_PROPERTY

PROPERTY PUBLIC FromBackStep : BOOL
GET
END_GET
END_PROPERTY

PROPERTY PUBLIC LastUsedKey : ULINT
GET
END_GET
END_PROPERTY

PROPERTY PUBLIC StepMemory_RO : I_ListOf_StepMemory_RO
GET
END_GET
END_PROPERTY

PROPERTY PUBLIC StepNumberHome : INT
GET
END_GET
END_PROPERTY

(*
Description
===========
| Condition to switch to the next step in automatic mode (also in manual mode if "ManualWithCondition" is TRUE) 
*)

PROPERTY PUBLIC Condition : BOOL
GET
END_GET
END_PROPERTY

PROPERTY PUBLIC DisableBackward : BOOL
GET
END_GET
END_PROPERTY

(*
Description
===========
| Step number to go to next
| 0 = subsequent step
*)
PROPERTY PUBLIC JumpAddress : INT
GET
END_GET
END_PROPERTY

(*
Description
===========
| If TRUE, property "Condition" is also active in manual mode
*)
PROPERTY PUBLIC ManualWithCondition : BOOL
GET
END_GET
END_PROPERTY

(*
Description
===========
| automatic: Control automatically jumps to the next step if Condition is TRUE
| manual: Input ManualForward must be pulsed TRUE to go to the next step
*)
PROPERTY PUBLIC mode : REFERENCE to T_processMode
GET
END_GET
END_PROPERTY

END_INTERFACE

// Step/processStep/I_processStep
INTERFACE I_processStep EXTENDS KOSTAL_AF2024_Core_System.I_Interface

(*
Description
===========
| Actual step number
*)
PROPERTY PUBLIC actual : INT
GET
END_GET
END_PROPERTY

METHOD PUBLIC CopyTo : BOOL
VAR_INPUT
	IN	:	I_processStep_CopyFrom;
END_VAR
END_METHOD

(*
Description
===========
| Requested step number (will be set with the next call of Header()
*)
PROPERTY PUBLIC request : INT
GET
END_GET
END_PROPERTY

(*
Description
===========
| Toggle signal for initialzation purposes
| Is set TRUE when Header() was called and the step number changed
| Is reset FALSE with the next call of Header() without changing step number
*)

PROPERTY PUBLIC toggle : BOOL
GET
END_GET
END_PROPERTY

END_INTERFACE

// Step/processStep/I_processStep_CopyFrom
INTERFACE I_processStep_CopyFrom EXTENDS KOSTAL_AF2024_Core_System.I_Interface

METHOD PUBLIC CopyFrom : BOOL
VAR_INPUT
	IN	: KOSTAL_AF2024_Core_System.I_Interface;
END_VAR
END_METHOD

END_INTERFACE

// Step/processStep_Control/StepMemory/ListOf/I_ListOf_StepMemory_RO
(*
	Read only Interface from List of DUT
*)
INTERFACE I_ListOf_StepMemory_RO EXTENDS KOSTAL_AF2024_Core_ListOf._I_Object_Base

METHOD PUBLIC CopyTo : BOOL
VAR_INPUT
	IN	: I_ListOf_StepMemory_CopyFrom;
END_VAR
END_METHOD

METHOD Get_I_RO : BOOL

VAR_INPUT
	Number		: UDINT;
	rFound_I	: REFERENCE TO I_T_StepMemory_RO;
	Response	: KOSTAL_AF2024_Core_functionResponse.I_T_functionResponse_Owner;
END_VAR
END_METHOD

PROPERTY PUBLIC MaxEntries : UDINT
GET
END_GET
END_PROPERTY

PROPERTY NumberOfMember : UDINT
GET
END_GET
END_PROPERTY

END_INTERFACE

// Step/processStep_Control/StepMemory/ListOf/I_ListOf_StepMemory_CopyFrom
(*
	The class implementing this interface can take over the contents from another instance with the same interface {I_DUT}.
	Typing takes place in the method.
*)
INTERFACE I_ListOf_StepMemory_CopyFrom EXTENDS KOSTAL_AF2024_Core_System.I_Interface

(*
	Copies the contents of another list {IN} into its own memory.
*)
METHOD PUBLIC CopyFrom : BOOL
VAR_INPUT
	IN	: KOSTAL_AF2024_Core_System.I_Interface;
END_VAR
END_METHOD

END_INTERFACE

// Step/processStep_Control/StepMemory/I_T_StepMemory_RO
INTERFACE I_T_StepMemory_RO EXTENDS KOSTAL_AF2024_Core_System.I_Interface

METHOD PUBLIC CopyTo : BOOL
VAR_INPUT
	IN	: I_T_StepMemory_CopyFrom;
END_VAR
END_METHOD

PROPERTY PUBLIC Actual : INT
GET
END_GET
END_PROPERTY

PROPERTY PUBLIC RegKey : ULINT
GET
END_GET
END_PROPERTY

PROPERTY PUBLIC Request : INT
GET
END_GET
END_PROPERTY

END_INTERFACE

// Step/processStep_Control/StepMemory/I_T_StepMemory_CopyFrom
INTERFACE I_T_StepMemory_CopyFrom EXTENDS KOSTAL_AF2024_Core_System.I_Interface

METHOD PUBLIC CopyFrom	:	BOOL
VAR_INPUT
	IN	: KOSTAL_AF2024_Core_System.I_Interface;
END_VAR
END_METHOD

END_INTERFACE

// Step/processStep_Control/I_ProcessStep_Control_Owner
INTERFACE I_ProcessStep_Control_Owner EXTENDS I_processStep_Owner

(*
Description
===========
| Select next step number dependent of Condition and JumpAddress
*)

METHOD PUBLIC Control : KOSTAL_AF2024_Core_functionResponse.T_functionResponse
END_METHOD

(*
Description
===========
| Apply changes in step sequence
| Call before the step sequence (see usage sample)
*)
METHOD PUBLIC Header
END_METHOD

//It is mandatory to link the parameters exclusively with pulses. 
METHOD PUBLIC LinkManual
VAR_INPUT
	Forward		: BOOL;	//Pulse one step forward in the step chain 
	Backward	: BOOL;	//Pulse one step backwards in the step chain
END_VAR
END_METHOD

(*
Description
===========
| Step change backward was successful - Use e.g. to reset requests
| Attention: Variable is reset with next call of Header()
*)
PROPERTY PUBLIC BackwardDone : BOOL
GET
END_GET
END_PROPERTY

(*
Description
===========
| Step change was successful - Use e.g. to reset requests
| Attention: Variable is reset with next call of Header()
*)
PROPERTY PUBLIC Done : BOOL
GET
END_GET
END_PROPERTY

PROPERTY PUBLIC FromBackStep : BOOL
GET
END_GET
END_PROPERTY

PROPERTY PUBLIC LastUsedKey : ULINT
GET
END_GET
END_PROPERTY

PROPERTY PUBLIC StepMemory : I_ListOf_StepMemory
GET
END_GET
END_PROPERTY

PROPERTY PUBLIC StepMemory_RO : I_ListOf_StepMemory_RO
GET
END_GET
END_PROPERTY

PROPERTY PUBLIC StepNumberHome : INT
GET
END_GET
SET
END_SET
END_PROPERTY

(*
Description
===========
| Condition to switch to the next step in automatic mode (also in manual mode if "ManualWithCondition" is TRUE) 
*)

PROPERTY PUBLIC Condition : BOOL
GET
END_GET
SET
END_SET
END_PROPERTY

PROPERTY PUBLIC DisableBackward : BOOL
GET
END_GET
SET
END_SET
END_PROPERTY

(*
Description
===========
| Step number to go to next
| 0 = subsequent step
*)
PROPERTY PUBLIC JumpAddress : INT
GET
END_GET
SET
END_SET
END_PROPERTY

(*
Description
===========
| If TRUE, property "Condition" is also active in manual mode
*)
PROPERTY PUBLIC ManualWithCondition : BOOL
GET
END_GET
SET
END_SET
END_PROPERTY

(*
Description
===========
| automatic: Control automatically jumps to the next step if Condition is TRUE
| manual: Input ManualForward must be pulsed TRUE to go to the next step
*)
PROPERTY PUBLIC mode : REFERENCE to T_processMode
GET
END_GET
SET
END_SET
END_PROPERTY

END_INTERFACE

// Step/processStep/I_processStep_Owner
INTERFACE I_processStep_Owner EXTENDS KOSTAL_AF2024_Core_System.I_Interface

(*
Description
===========
| Actual step number
*)
PROPERTY PUBLIC actual : INT
GET
END_GET
END_PROPERTY

METHOD PUBLIC clear
END_METHOD

METHOD PUBLIC CopyFrom : BOOL
VAR_INPUT
	IN	: KOSTAL_AF2024_Core_System.I_Interface;
END_VAR
END_METHOD

METHOD PUBLIC CopyTo : BOOL
VAR_INPUT
	IN	:	I_processStep_CopyFrom;
END_VAR
END_METHOD

(*
Description
===========
| Decrease step number by one (will be set with the next call of Header()
*)
METHOD DEC : KOSTAL_AF2024_Core_functionResponse.T_functionResponse
VAR_INPUT
END_VAR
END_METHOD

(*
Description
===========
| Apply changes in step sequence
| Call before or after the step sequence (see usage sample)
*)
METHOD PUBLIC Header
VAR_INPUT
END_VAR
END_METHOD

(*
Description
===========
| Increase step number by one (will be set with the next call of Header()
*)
METHOD INC : KOSTAL_AF2024_Core_functionResponse.T_functionResponse
END_METHOD

(*
Description
===========
| Reset step sequence to 0
*)
METHOD PUBLIC init
END_METHOD

(*
Description
===========
| Requested step number (will be set with the next call of Header()
*)
PROPERTY PUBLIC request : INT
GET
END_GET
END_PROPERTY

(*
Description
===========
| Select step number (will be set with the next call of Header()
| Same function as property request
| Parameters:
| 	request: INT - step number to go to
*)
METHOD PUBLIC set

VAR_INPUT
	request	: INT;	//INT
END_VAR
END_METHOD

(*
Description
===========
| Toggle signal for initialzation purposes
| Is set TRUE when Header() was called and the step number changed
| Is reset FALSE with the next call of Header() without changing step number
*)

PROPERTY PUBLIC toggle : BOOL
GET
END_GET
END_PROPERTY

END_INTERFACE

// Step/processStep_Control/StepMemory/ListOf/I_ListOf_StepMemory
(*
	Full qualified access Interface from List of DUT
*)
INTERFACE I_ListOf_StepMemory EXTENDS KOSTAL_AF2024_Core_ListOf._I_Object_Base_Owner

//Add a new instance of FB_Dut and copy content from [IN] to the new instance
METHOD PUBLIC Add_DUT : BOOL
VAR_INPUT
	IN				: KOSTAL_AF2024_Core_System.I_Interface;
	Response	: KOSTAL_AF2024_Core_functionResponse.I_T_functionResponse_Owner;
END_VAR
END_METHOD

METHOD Clear
VAR_INPUT
END_VAR
END_METHOD

METHOD PUBLIC CopyFrom : BOOL
VAR_INPUT
	IN	: KOSTAL_AF2024_Core_System.I_Interface;
END_VAR
END_METHOD

METHOD PUBLIC CopyTo : BOOL
VAR_INPUT
	IN	: I_ListOf_StepMemory_CopyFrom;
END_VAR
END_METHOD

METHOD PUBLIC Delete_DUT : BOOL
VAR_INPUT
	Number	: UDINT;	//Number of DUT in List
	Response	: KOSTAL_AF2024_Core_functionResponse.I_T_functionResponse_Owner;
END_VAR
END_METHOD

//Get full access to content 
METHOD Get_I : BOOL

VAR_INPUT
	Number		: UDINT;
	rFound_I	: REFERENCE TO I_T_StepMemory;
	Response	: KOSTAL_AF2024_Core_functionResponse.I_T_functionResponse_Owner;
END_VAR
END_METHOD

METHOD Get_I_RO : BOOL

VAR_INPUT
	Number		: UDINT;
	rFound_I	: REFERENCE TO I_T_StepMemory_RO;
	Response	: KOSTAL_AF2024_Core_functionResponse.I_T_functionResponse_Owner;
END_VAR
END_METHOD

PROPERTY PUBLIC MaxEntries : UDINT
GET
END_GET
SET
END_SET
END_PROPERTY

PROPERTY NumberOfMember : UDINT
GET
END_GET
END_PROPERTY

END_INTERFACE

// Step/processStep_Control/StepMemory/I_T_StepMemory
INTERFACE I_T_StepMemory EXTENDS I_T_StepMemory_RO

METHOD PUBLIC Clear
END_METHOD

METHOD PUBLIC CopyFrom	:	BOOL
VAR_INPUT
	IN	: KOSTAL_AF2024_Core_System.I_Interface;
END_VAR
END_METHOD

PROPERTY PUBLIC Actual : INT
SET
END_SET
END_PROPERTY

PROPERTY PUBLIC RegKey : ULINT
SET
END_SET
END_PROPERTY

PROPERTY PUBLIC Request : INT
GET
END_GET
SET
END_SET
END_PROPERTY

END_INTERFACE

// Step/processStep_Control/StepMemory/ListOf/FB_ListOf_T_StepMemory
(*
	A template for creating a list of typed classes (FBs)
*)
FUNCTION_BLOCK FB_ListOf_T_StepMemory EXTENDS KOSTAL_AF2024_Core_ListOf._FB_Object_Base  IMPLEMENTS I_ListOf_StepMemory_RO, I_ListOf_StepMemory_CopyFrom, I_ListOf_StepMemory

VAR
	//Use the {_Dummy} to ensure that a valid interface is always returned.
	_Dummy			: T_StepMemory;
	_MaxEntries	: UDINT:= UDINT#128;
END_VAR

(*
	Returns the typed owner interface in the reference variable.
	In the event of an error, the return value becomes FALSE and the interface refers to the {_Dummy}.
*)
METHOD PROTECTED _get_I : BOOL

VAR_INPUT
	Member		: KOSTAL_AF2024_Core_System.I_Interface;
	rFound_I	: REFERENCE TO I_T_StepMemory;
	rResult		: KOSTAL_AF2024_Core_functionResponse.I_T_functionResponse_Owner;
END_VAR

VAR
	_iObj			: I_T_StepMemory;
	_Success	: BOOL;
END_VAR

IF NOT SUPER^._verifyMember(Member, rResult)	THEN 
	IF __ISVALIDREF(rFound_I)	THEN	rFound_I:= _Dummy;	END_IF
	RETURN;	
END_IF

_Success:= __QUERYINTERFACE(Member, _iObj);

//return dummy if no valid DUT is found
IF NOT _Success OR (_iObj = 0)	THEN	

	IF __ISVALIDREF(rFound_I)	THEN	rFound_I:= _Dummy;	END_IF	
	IF rResult <> 0						THEN	rResult.success:= FALSE;	
																	rResult.status:= "__QueryInterface failed - return Dummy";	
	END_IF	

	RETURN;	

END_IF

IF __ISVALIDREF(rFound_I)	THEN	rFound_I:= _iObj;	END_IF
IF rResult <> 0						THEN	rResult.success:= TRUE;
																rResult.status:= "Successful";
END_IF

_get_I:= TRUE;
END_METHOD

(*
	Returns the typed interface in the reference variable.
	In the event of an error, the return value becomes FALSE and the interface refers to the {_Dummy}.
*)
METHOD PROTECTED _get_I_RO : BOOL

VAR_INPUT
	Member		: KOSTAL_AF2024_Core_System.I_Interface;
	rFound_I	: REFERENCE TO I_T_StepMemory_RO;
	rResult		: KOSTAL_AF2024_Core_functionResponse.I_T_functionResponse_Owner;
END_VAR

VAR
	_iObj	: I_T_StepMemory_RO;
	_Success: BOOL;
END_VAR

IF NOT SUPER^._verifyMember(Member, rResult)	THEN 
	IF __ISVALIDREF(rFound_I)	THEN	rFound_I:= _Dummy;	END_IF
	RETURN;	
END_IF

_Success:= __QUERYINTERFACE(Member, _iObj);

//return dummy if no valid DUT is found
IF NOT _Success OR (_iObj = 0)	THEN	

	IF __ISVALIDREF(rFound_I)	THEN	rFound_I:= _Dummy;	END_IF	
	IF rResult <> 0						THEN	rResult.success:= FALSE;		
																	rResult.status:= "__QueryInterface failed - return Dummy";	
	END_IF	

	RETURN;	

END_IF

IF __ISVALIDREF(rFound_I)	THEN	rFound_I:= _iObj;	END_IF
IF rResult <> 0						THEN	rResult.success:= TRUE;
																rResult.status:= "Successful";
END_IF

_get_I_RO:= TRUE;
END_METHOD

(*
	Cleans the custom class {FB_DUT} and removes it from memory.
*)
METHOD PROTECTED  _removePayLoad : BOOL
VAR_INPUT
	Member	: KOSTAL_AF2024_Core_System.I_Interface;
	Result	: KOSTAL_AF2024_Core_functionResponse.I_T_functionResponse_Owner;
END_VAR

VAR
	_iObj			: I_T_StepMemory;
	_pFB_DUT	:	POINTER TO T_StepMemory;
	_Success	: BOOL;
END_VAR


IF NOT SUPER^._removePayload(Member, Result)	THEN RETURN;	END_IF

_Success:= __QUERYINTERFACE(Member, _iObj);

IF NOT _Success	THEN	RETURN;	END_IF
IF _iObj = 0		THEN	RETURN;	END_IF

_iObj.Clear();

_Success  := __QUERYPOINTER(_iObj, _pFB_DUT);

IF NOT _Success	THEN	RETURN;	END_IF
IF _pFB_DUT = 0	THEN	RETURN;	END_IF

__DELETE(_pFB_DUT);
END_METHOD

(*
	Overload the method from the base class to verify the custom interface. 
	The local method {_get_I_Owner()} is used for this.
*)
METHOD PROTECTED _verifyMember : BOOL
VAR_INPUT
	Member	: KOSTAL_AF2024_Core_System.I_Interface;
	Result	: KOSTAL_AF2024_Core_functionResponse.I_T_functionResponse_Owner;
END_VAR


_verifyMember:= _get_I(Member, 0, Result);
END_METHOD

(*
	Add a new instance of FB_Dut and copy content from [IN] to the new instance
*)
METHOD PUBLIC Add_DUT : BOOL
VAR_INPUT
	IN				: KOSTAL_AF2024_Core_System.I_Interface;
	Response	: KOSTAL_AF2024_Core_functionResponse.I_T_functionResponse_Owner;
END_VAR

VAR
	_pDUT: POINTER TO T_StepMemory;
	_response: KOSTAL_AF2024_Core_functionResponse.T_functionResponse;
END_VAR

_response.clear();

IF _Count	> _MaxEntries THEN 
	IF Response <> 0 THEN	Response.success:= FALSE;	Response.status:= "Max entries overflow";	END_IF
	RETURN;	
END_IF

_pDUT:= __NEW(T_StepMemory);

IF _pDUT = 0 THEN
	_response.status:= "cannot create new object";
	IF Response <> 0 THEN	Response.CopyFrom(_response);	END_IF
	RETURN;
END_IF

IF NOT _pDUT^.CopyFrom(IN) THEN
	Response.success:= FALSE;	Response.status:= "cannot copy content";
	__DELETE(_pDUT);
	RETURN;
END_IF

SUPER^._addMember(_pDUT^, _response);

_pDUT^.RegKey:= _RegKeyValue;

IF Response <> 0 THEN	Response.CopyFrom(_response);	END_IF

Add_DUT:= _response.success;
END_METHOD

(*
	Makes the protected method public.
*)
METHOD Clear

SUPER^._clear();
END_METHOD

(*
	Copies the contents of another list {IN} into its own memory.
*)
METHOD PUBLIC CopyFrom : BOOL
VAR_INPUT
	IN	: KOSTAL_AF2024_Core_System.I_Interface;
END_VAR

VAR
	_udi		: UDINT;

	_obj		: I_ListOf_StepMemory_RO;
	_IDUT		: I_T_StepMemory_RO;

	_obj2		: I_ListOf_StepMemory;
	_IDUT2	: I_T_StepMemory;

	_bFound	:	BOOL;
END_VAR
IF IN = 0 THEN RETURN;	END_IF

_clear();

_bFound:= __QUERYINTERFACE(IN, _obj);

IF _bFound AND_THEN _obj <> 0 THEN
	
	FOR _udi:= 1 TO _obj.NumberOfMember DO
		IF _obj.Get_I_RO(_udi, _IDUT, 0)	THEN	Add_DUT(_IDUT, 0);	END_IF
	END_FOR

	CopyFrom:= TRUE;

	RETURN;	

END_IF


_bFound:= __QUERYINTERFACE(IN, _obj2);

IF _bFound AND_THEN _obj2 <> 0 THEN
	
	FOR _udi:= 1 TO _obj2.NumberOfMember DO
		IF _obj2.Get_I(_udi, _IDUT2, 0)	THEN	Add_DUT(_IDUT2, 0);	END_IF
	END_FOR

	CopyFrom:= TRUE;

	RETURN;	

END_IF
END_METHOD

(*
	Copies the own content into another list created at the parameter {IN}.
*)
METHOD PUBLIC CopyTo : BOOL
VAR_INPUT
	IN	: I_ListOf_StepMemory_CopyFrom;
END_VAR

IF IN = 0 THEN RETURN;	END_IF

CopyTo:= IN.CopyFrom(THIS^);
END_METHOD

(*
	Deletes the class specified with the {Number} from the list.
*)
METHOD PUBLIC Delete_DUT : BOOL
VAR_INPUT
	Number		: UDINT;	//Number of DUT in List
	Response	: KOSTAL_AF2024_Core_functionResponse.I_T_functionResponse_Owner;
END_VAR

VAR
	_response	: KOSTAL_AF2024_Core_functionResponse.T_functionResponse;
	_Success	: BOOL;
	_Member		: KOSTAL_AF2024_Core_System.I_Interface;
END_VAR

IF Number = 0 THEN
	_response.clear(); _response.status:= "Number is out of range (1..n)"; 
	IF Response <> 0 THEN	Response.CopyFrom(_response);	END_IF
	RETURN;
END_IF

Delete_DUT:= SUPER^._removeMemberByIndex(Number - 1, _response);

IF Response <> 0 THEN	Response.CopyFrom(_response);	END_IF

Delete_DUT:= _response.success;
END_METHOD

(*
	Get full access to content of Member with {Number}
*) 
METHOD Get_I : BOOL

VAR_INPUT
	Number		: UDINT;
	rFound_I	: REFERENCE TO I_T_StepMemory;
	Response	: KOSTAL_AF2024_Core_functionResponse.I_T_functionResponse_Owner;
END_VAR

VAR
	_Member				: KOSTAL_AF2024_Core_System.I_Interface;
	_response			: KOSTAL_AF2024_Core_functionResponse.T_functionResponse;
END_VAR
IF Number = 0 THEN
	IF __ISVALIDREF(rFound_I)	THEN	rFound_I:= _Dummy;	END_IF
	_response.clear(); _response.status:= "Number is out of range (1..n)"; 
	IF Response <> 0 THEN	Response.CopyFrom(_response);	END_IF
	RETURN;
END_IF

IF NOT SUPER^._findMemberByIndex(Number - 1, _Member, Response) THEN

 IF __ISVALIDREF(rFound_I) THEN	rFound_I:= _Dummy;	END_IF

ELSE

	Get_I:= _get_I(_Member, rFound_I, Response);
	
END_IF
END_METHOD

(*
	Get readonly access to content of Member with {Number}
*) 
METHOD Get_I_RO : BOOL

VAR_INPUT
	Number		: UDINT;
	rFound_I	: REFERENCE TO I_T_StepMemory_RO;
	Response	: KOSTAL_AF2024_Core_functionResponse.I_T_functionResponse_Owner;
END_VAR

VAR
	_Member		: KOSTAL_AF2024_Core_System.I_Interface;
	_response	: KOSTAL_AF2024_Core_functionResponse.T_functionResponse;
END_VAR
IF Number = 0 THEN
	IF __ISVALIDREF(rFound_I)	THEN	rFound_I:= _Dummy;	END_IF
	_response.clear(); _response.status:= "Number is out of range (1..n)"; 
	IF Response <> 0 THEN	Response.CopyFrom(_response);	END_IF
	RETURN;
END_IF

IF NOT SUPER^._findMemberByIndex(Number - 1, _Member, Response) THEN

 IF __ISVALIDREF(rFound_I) THEN	rFound_I:= _Dummy;	END_IF

ELSE

	Get_I_RO:= _get_I_RO(_Member, rFound_I, Response);
	
END_IF
END_METHOD

PROPERTY PUBLIC MaxEntries : UDINT
GET

MaxEntries:= _MaxEntries;
END_GET
SET

_MaxEntries:= MaxEntries;
END_SET
END_PROPERTY

(*
	Number of Member in list.
*)
PROPERTY NumberOfMember : UDINT
GET

NumberOfMember:= SUPER^._NumberOfMember;
END_GET
END_PROPERTY

END_FUNCTION_BLOCK

// Step/processStep_Control/StepMemory/T_StepMemory
{attribute 'enable_dynamic_creation'}
FUNCTION_BLOCK PUBLIC T_StepMemory IMPLEMENTS I_T_StepMemory_RO, I_T_StepMemory, I_T_StepMemory_CopyFrom
VAR
	_Actual		: INT;	//Contains the actual step
	_Request	: INT;	//Contains the requested step
	_RegKey		: ULINT:= ULINT#0;	//Handled exclusively in this class  
END_VAR

METHOD PUBLIC Clear

_Actual		:= INT#0;
_Request	:= INT#0;
_RegKey		:= ULINT#0;
END_METHOD

METHOD PUBLIC CopyFrom	:	BOOL
VAR_INPUT
	IN	: KOSTAL_AF2024_Core_System.I_Interface;
END_VAR

VAR
	_obj		: I_T_StepMemory_RO;
	_obj2		: I_T_StepMemory;
	_bFound	:	BOOL;
END_VAR

IF IN = 0 THEN RETURN;	END_IF

Clear();

_bFound:= __QUERYINTERFACE(IN, _obj);

IF _bFound AND_THEN _obj <> 0 THEN

	_Actual		:= _obj.Actual;
	_Request	:= _obj.Request;
	_RegKey		:= _obj.RegKey;
	
	CopyFrom:= TRUE;
	
	RETURN;	

END_IF

_bFound:= __QUERYINTERFACE(IN, _obj2);

IF _bFound AND_THEN _obj2 <> 0 THEN

	_Actual		:= _obj2.Actual;
	_Request	:= _obj2.Request;
	_RegKey		:= _obj2.RegKey;
	
	CopyFrom:= TRUE;
	
	RETURN;	

END_IF
END_METHOD

METHOD PUBLIC CopyTo : BOOL
VAR_INPUT
	IN	: I_T_StepMemory_CopyFrom;
END_VAR

IF IN = 0 THEN RETURN;	END_IF

CopyTo:= IN.CopyFrom(THIS^);
END_METHOD

PROPERTY PUBLIC Actual : INT
GET

Actual:= _Actual;
END_GET
SET

_Actual:= Actual;
END_SET
END_PROPERTY

PROPERTY PUBLIC RegKey : ULINT
GET

RegKey:= _RegKey;
END_GET
SET

_RegKey:= RegKey;
END_SET
END_PROPERTY

PROPERTY PUBLIC Request : INT
GET

Request:= _Request;
END_GET
SET

_Request:= Request;
END_SET
END_PROPERTY

END_FUNCTION_BLOCK

// Step/processStep_Flow/FB_processStep_Flow
(*

:Author: Frank Dümpelmann <f.duempelmann@kostal.com>
:Date: 2019-03-29

Function
========
| Extends FB_processStep

Methods and Properties
======================
| See bottom of this document for a detailed description of each method or property
*)

{attribute 'enable_dynamic_creation'}
FUNCTION_BLOCK PUBLIC FB_processStep_Flow EXTENDS FB_processStep IMPLEMENTS I_processStep_Flow, I_processStep_Flow_Owner

VAR
	_Found	: BOOL;
END_VAR

METHOD PUBLIC clear

_Found:= FALSE;

SUPER^.clear();
END_METHOD

(*
Description
===========
| Apply changes in step sequence
| Call before or after the step sequence (see usage sample)
*)
METHOD PUBLIC Header
VAR_INPUT
END_VAR

_Found:= FALSE;
END_METHOD

(*
Description
===========
| Reset step sequence to 0
*)
METHOD PUBLIC init

_Found:= FALSE;

SUPER^.init();
END_METHOD

(*
| Description
| ============
| Returns TRUE if step.active is equal stepNumber 
*)

METHOD PUBLIC isActive : BOOL
VAR_INPUT
	stepNumber	: INT;
END_VAR
 
isActive:= _request = stepNumber;

IF NOT isActive THEN RETURN;	END_IF

_Found:= TRUE;

SUPER^.Header();
END_METHOD

METHOD PUBLIC isCalledExternally : BOOL
VAR_INPUT
END_VAR

isCalledExternally:= _actual <> _request;
END_METHOD

METHOD PUBLIC NotFound : BOOL
VAR_INPUT
END_VAR

NotFound:= NOT _Found;
END_METHOD

END_FUNCTION_BLOCK

// Step/processStep_Flow/I_processStep_Flow
INTERFACE I_processStep_Flow EXTENDS I_processStep

METHOD PUBLIC isCalledExternally : BOOL
VAR_INPUT
END_VAR
END_METHOD

METHOD PUBLIC NotFound : BOOL
VAR_INPUT
END_VAR
END_METHOD

END_INTERFACE

// Step/processStep_Flow/I_processStep_Flow_Owner
INTERFACE I_processStep_Flow_Owner EXTENDS I_processStep_Owner

METHOD PUBLIC clear
END_METHOD

(*
Description
===========
| Apply changes in step sequence
| Call before or after the step sequence (see usage sample)
*)
METHOD PUBLIC Header
VAR_INPUT
END_VAR
END_METHOD

(*
Description
===========
| Reset step sequence to 0
*)
METHOD PUBLIC init
END_METHOD

(*
| Description
| ============
| Returns TRUE if step.active is equal stepNumber 
*)

METHOD PUBLIC isActive : BOOL
VAR_INPUT
	stepNumber	: INT;
END_VAR
END_METHOD

METHOD PUBLIC isCalledExternally : BOOL
VAR_INPUT
END_VAR
END_METHOD

METHOD PUBLIC NotFound : BOOL
VAR_INPUT
END_VAR
END_METHOD

END_INTERFACE
